(* IEC 61131-3 sources: Test-Git_ESME26/TestProgettoESME_26.fbsproj/PacDriveLib Migration/Motion/Homing, 18 files *)

(* ---- PDL_FC_ReadDriveEncoder.fn.st ---- *)
FUNCTION PDL_FC_ReadDriveEncoder: BOOL
VAR_INPUT
	i_ifDrive			: MOIN.IF_Axis;
	i_lrHomePos			: LREAL;
	i_lrAbsEncOffset	: LREAL;
	i_lrUserPeriod		: LREAL;
END_VAR
VAR_OUTPUT
	q_etDiag			: GD.ET_Diag := GD.ET_Diag.OK;
	q_etDiagExt			: PDL_ET_DiagExt := PDL_ET_DiagExt.OK;
	q_sMsg				: STRING[80];
END_VAR
VAR
	ifGetParentDevice   : DTSI.IF_GetParentDevice;
	ifDeviceAccess		: DTSI.IF_DeviceAccess;
	ifEncoderAccess		: DDI.IF_EncoderAccess;
	ifEncoder			: DDI.IF_Encoder;
	ifScalingAccess     : DMFI.IF_ScalingAccess;
	ifScaling		    : DMFI.IF_Scaling;
	xSuccess			: BOOL;
	lrEncoderPeriode:	LREAL;
	lrEncPosition:		LREAL;
	lrModuloPosition:	LREAL;
	lrHomePosition:		LREAL;
	lrTurns:			LREAL;
	lrEncoderRange:		LREAL;
	fbSetPos			: PLCO.MC_SetPosition;
END_VAR
VAR CONSTANT
	c_lrRealNull				: LREAL := 10E-12;
END_VAR

IF i_ifDrive = 0 THEN
	q_etDiag	:= GD.ET_Diag.InputParameterInvalid;
	q_etDiagExt := PDL_ET_DiagExt.DriveInvalid;
	q_sMsg		:= 'i_ifDrive - Invalid Interface';
	RETURN;
END_IF

xSuccess := __QUERYINTERFACE(i_ifDrive, ifGetParentDevice);
IF NOT xSuccess OR ifGetParentDevice = 0 THEN
	q_etDiag	:= GD.ET_Diag.InputParameterInvalid;
	q_etDiagExt := PDL_ET_DiagExt.DriveInvalid;
	q_sMsg		:= 'i_ifDrive - IF_GetParentDevice not implemented.';
	RETURN;
END_IF
ifDeviceAccess := ifGetParentDevice.GetParentDevice();

xSuccess := __QUERYINTERFACE(ifDeviceAccess,ifEncoderAccess );
IF (NOT xSuccess OR ifEncoderAccess = 0) THEN
	q_etDiag	:= GD.ET_Diag.InputParameterInvalid;
	q_etDiagExt := PDL_ET_DiagExt.DriveInvalid;
	q_sMsg		:= 'i_ifDrive - IF_Encoder not implemented.';
	RETURN;
END_IF
ifEncoder := ifEncoderAccess.Encoder;

xSuccess := __QUERYINTERFACE(ifDeviceAccess,ifScalingAccess );
IF (NOT xSuccess OR ifScalingAccess = 0) THEN
	q_etDiag	:= GD.ET_Diag.InputParameterInvalid;
	q_etDiagExt := PDL_ET_DiagExt.DriveInvalid;
	q_sMsg		:= 'i_ifDrive - IF_Scaling not implemented.';
	RETURN;
END_IF
ifScaling := ifScalingAccess.Scaling;
// Allgemeine Berehcnung ohne unterscheidung des Gebertyps			30.09.2009/ck
lrEncoderRange := ifEncoder.Revolutions;
IF (ABS(lrEncoderRange) < 1.0E-3) THEN
	q_etDiag	:= GD.ET_Diag.DriveConditionInvalid;
	q_etDiagExt := PDL_ET_DiagExt.DriveEncoderInvalid;
	q_sMsg		:= '';
	RETURN;
ELSE
	lrEncoderPeriode := lrEncoderRange * ifScaling.PositionResolution * TO_LREAL(ifScaling.GearIn) / TO_LREAL(ifScaling.GearOut);
END_IF

IF (i_lrUserPeriod < 0.0) THEN
	q_etDiag	:= GD.ET_Diag.InputParameterInvalid;
	q_etDiagExt := PDL_ET_DiagExt.UserPeriodRange;
	q_sMsg		:= '0.0 <= i_lrUserPeriod';

ELSIF (i_lrUserPeriod < c_lrRealNull) AND
	( (i_lrAbsEncOffset < c_lrRealNull) OR (i_lrAbsEncOffset > (lrEncoderPeriode - c_lrRealNull)) ) THEN
	q_etDiag	:= GD.ET_Diag.InputParameterInvalid;
	q_etDiagExt := PDL_ET_DiagExt.AbsEncOffsetRange;
	q_sMsg		:= STANDARD.CONCAT('0.0 < i_lrAbsEncOffset <= ', SE_CTBX.FC_LrealToString(i_sFormat := '#0.00', i_lrInput := lrEncoderPeriode - c_lrRealNull));

(* Check if UserPeriode fits into EncoderPeriode *)
ELSIF(i_lrUserPeriod > c_lrRealNull) AND
		(ABS(lrEncoderPeriode/i_lrUserPeriod - TRUNC_INT(lrEncoderPeriode / i_lrUserPeriod)) > c_lrRealNull ) THEN
	q_etDiag	:= GD.ET_Diag.InputParameterInvalid;
	q_etDiagExt := PDL_ET_DiagExt.UserPeriodRange;
	q_sMsg		:= STANDARD.CONCAT('i_lrUserPeriod has to be a divsior of ', SE_CTBX.FC_LrealToString(i_sFormat := '#0.00', i_lrInput := lrEncoderPeriode));

ELSE

	IF NOT ifScaling.InvertDirection THEN				(* motor direction right (true) *)
		lrEncPosition := ifEncoder.Position;
	ELSE
		lrEncPosition := lrEncoderPeriode - ifEncoder.Position;
	END_IF

(* In a round axis, position is always within the user period *)
	IF i_lrUserPeriod > c_lrRealNull THEN
		lrHomePosition := i_lrHomePos + lrEncPosition - lrEncoderPeriode/2.0;

		lrTurns :=  TRUNC_INT(lrHomePosition / i_lrUserPeriod);
		IF lrHomePosition < 0 THEN
			lrTurns := lrTurns - 1;
		END_IF

		lrModuloPosition := lrHomePosition - lrTurns * i_lrUserPeriod;

	ELSE
		lrModuloPosition := i_lrHomePos + lrEncPosition - i_lrAbsEncOffset;
	END_IF

	fbSetPos(Axis := i_ifDrive, Position := lrModuloPosition, Relative := FALSE, Execute := TRUE);

	IF fbSetPos.Error THEN
		q_etDiag	:= GD.ET_Diag.UnexpectedProgramBehavior;
		q_etDiagExt := PDL_ET_DiagExt.UnexpectedDiagExt;
		q_sMsg		:= CONCAT('Setpos: ', TO_STRING(fbSetPos.ErrorId));
	END_IF
END_IF

(* ---- PDL_FC_RestoreAxisPosition.fn.st ---- *)
FUNCTION PDL_FC_RestoreAxisPosition : BOOL
VAR_INPUT
	i_ifDrive           : MOIN.IF_Axis;
	i_lrUserPeriod      : LREAL;
	i_lrRestoreWindow   : LREAL;
	i_stRestorePosition : PDL_ST_AxisRestorePosition;
END_VAR
VAR_OUTPUT
	q_etDiag    : GD.ET_Diag     := GD.ET_Diag.OK;
	q_etDiagExt : PDL_ET_DiagExt := PDL_ET_DiagExt.OK;
	q_sMsg      : STRING[80];
END_VAR
VAR
	xSuccess            : BOOL;
	lrEncMaxPos         : LREAL;
	lrEncDiff           : LREAL;
	lrCalcAxisPos       : LREAL;
	dinPeriode          : DINT;
	diSercosState       : DINT;
	lrEncPos            : LREAL;
	lrAxisPosition      : LREAL;
	lrEncPosition       : LREAL;
	lrCheckSum          : LREAL;
	lrAxisEncPosition   : LREAL;
	lrAxisEncPosition2  : LREAL;
	diAxisGearIn        : DINT;
	diAxisGearOut       : DINT;
	lrAxisFeedConstant  : LREAL;
	diCount             : DINT;
	lrEncoderRange      : LREAL;
	ifScalingAccess     : DMFI.IF_ScalingAccess;
	ifScaling           : DMFI.IF_Scaling;
	ifGetParentDevice   : DTSI.IF_GetParentDevice;
	ifDeviceAccess      : DTSI.IF_DeviceAccess;
	ifEncoderAccess     : DDI.IF_EncoderAccess;
	ifEncoder           : DDI.IF_Encoder;
	fbSetPos            : PLCO.MC_SetPosition;
	xAxisDirection      : BOOL;

END_VAR
VAR CONSTANT
	c_lrDelta : LREAL := 0.01;
END_VAR

IF i_ifDrive = 0 THEN
	q_etDiag	:= GD.ET_Diag.InputParameterInvalid;
	q_etDiagExt := PDL_ET_DiagExt.DriveInvalid;
	q_sMsg		:= 'i_ifDrive - Invalid Interface';
	RETURN;
END_IF

xSuccess := __QUERYINTERFACE(i_ifDrive, ifGetParentDevice);
IF NOT xSuccess OR ifGetParentDevice = 0 THEN
	q_etDiag	:= GD.ET_Diag.InputParameterInvalid;
	q_etDiagExt := PDL_ET_DiagExt.DriveInvalid;
	q_sMsg		:= 'i_ifDrive - IF_GetParentDevice not implemented.';
	RETURN;
END_IF

ifDeviceAccess := ifGetParentDevice.GetParentDevice();

xSuccess := __QUERYINTERFACE(ifDeviceAccess,ifScalingAccess );
IF (NOT xSuccess OR ifScalingAccess = 0) THEN
	q_etDiag	:= GD.ET_Diag.InputParameterInvalid;
	q_etDiagExt := PDL_ET_DiagExt.DriveInvalid;
	q_sMsg		:= 'i_ifDrive - IF_Scaling not implemented.';
	RETURN;
END_IF
ifScaling := ifScalingAccess.Scaling;

xSuccess := __QUERYINTERFACE(ifDeviceAccess,ifEncoderAccess );
IF (NOT xSuccess OR ifEncoderAccess = 0) THEN
	q_etDiag	:= GD.ET_Diag.InputParameterInvalid;
	q_etDiagExt := PDL_ET_DiagExt.DriveInvalid;
	q_sMsg		:= 'i_ifDrive - IF_Encoder not implemented.';
	RETURN;
END_IF
ifEncoder := ifEncoderAccess.Encoder;

(*--------------------------------------------------------------------------------------------------------------------------------------------------*)
(* read values *)
(*--------------------------------------------------------------------------------------------------------------------------------------------------*)
	lrAxisPosition := i_stRestorePosition.lrAxisPosition;
	lrEncPosition := i_stRestorePosition.lrEncPosition;
	lrCheckSum := i_stRestorePosition.lrCheckSum;

	IF (((lrAxisPosition + lrEncPosition + c_lrDelta) < lrCheckSum) OR
		((lrAxisPosition + lrEncPosition - c_lrDelta) > lrCheckSum)) THEN

		q_etDiag	:= GD.ET_Diag.InputParameterInvalid;
		q_etDiagExt := PDL_ET_DiagExt.CheckSumInvalid;
		q_sMsg		:= '';
		RETURN;
	END_IF

(*--------------------------------------------------------------------------------------------------------------------------------------------------*)
(* Check Sercos state and read values *)
(*--------------------------------------------------------------------------------------------------------------------------------------------------*)
FOR diCount := 1 TO 3 DO

	diSercosState := FC_GetSercosState();
	IF diSercosState = 4 THEN
		lrAxisEncPosition := ifEncoder.Position;
		diAxisGearIn := TO_DINT(ifScaling.GearIn);
		diAxisGearOut := TO_DINT(ifScaling.GearOut);
		lrAxisFeedConstant := ifScaling.PositionResolution;
		xAxisDirection := NOT ifScaling.InvertDirection;
	ELSE
		q_etDiag	:= GD.ET_Diag.SercosConditionInvalid;
		q_etDiagExt := PDL_ET_DiagExt.SercosNotInPhaseFour;
		q_sMsg		:= '';
		RETURN;
	END_IF

(*--------------------------------------------------------------------------------------------------------------------------------------------------*)
(* Berechnung der maximale Encoder Position *)
(*--------------------------------------------------------------------------------------------------------------------------------------------------*)

	// Allgemeine Berechnung ohne Unterscheidung des Gebertyps
	lrEncoderRange := ifEncoder.Revolutions;
	IF (ABS(lrEncoderRange) < 1.0E-3) THEN
		q_etDiag	:= GD.ET_Diag.DriveConditionInvalid;
		q_etDiagExt := PDL_ET_DiagExt.DriveEncoderInvalid;
		q_sMsg		:= '';
		RETURN;
	ELSE
		lrEncMaxPos := lrEncoderRange * lrAxisFeedConstant * TO_LREAL(diAxisGearIn) / TO_LREAL(diAxisGearOut);
	END_IF

(*--------------------------------------------------------------------------------------------------------------------------------------------------*)
(* Differenz der Geberposition *)
(*--------------------------------------------------------------------------------------------------------------------------------------------------*)
	IF xAxisDirection THEN		(* +++ Rechtslauf +++ *)
		lrEncDiff := lrAxisEncPosition - lrEncPosition;
		IF lrEncDiff > lrEncMaxPos/2 THEN
			lrEncPos := lrAxisEncPosition - lrEncMaxPos;
			lrEncDiff := lrEncDiff - lrEncMaxPos;
		ELSIF lrEncDiff < -lrEncMaxPos/2 THEN
			lrEncPos := lrAxisEncPosition + lrEncMaxPos;
			lrEncDiff := lrEncDiff + lrEncMaxPos ;
		ELSE
			lrEncPos := lrAxisEncPosition;
		END_IF
		lrCalcAxisPos := lrEncPos - lrEncPosition + lrAxisPosition;

	ELSE						(* +++ Linkslauf +++ *)
		lrEncDiff:=  lrEncPosition - lrAxisEncPosition;	(*  lrEncMaxPos - lrAxisEncPosition
																 - (lrEncMaxPos- lrEncPos_Retain) *)
		IF lrEncDiff > lrEncMaxPos/2 THEN
			lrEncPos :=  - lrAxisEncPosition;				(* lrEncMaxPos - lrAxisEncPosition - lrEncMaxPos *)
			lrEncDiff := lrEncDiff - lrEncMaxPos;
		ELSIF lrEncDiff < -lrEncMaxPos/2 THEN
			lrEncPos := 2*lrEncMaxPos - lrAxisEncPosition;	(* lrEncMaxPos - lrAxisEncPosition + lrEncMaxPos *)
			lrEncDiff := lrEncDiff + lrEncMaxPos ;
		ELSE
			lrEncPos := lrEncMaxPos - lrAxisEncPosition;
		END_IF
		lrCalcAxisPos := lrEncPos -  (lrEncMaxPos - lrEncPosition) + lrAxisPosition;
	END_IF

(*--------------------------------------------------------------------------------------------------------------------------------------------------*)
(* check if in Window *)
(*--------------------------------------------------------------------------------------------------------------------------------------------------*)
	IF ABS(lrEncDiff) > ABS(i_lrRestoreWindow) THEN	(* Maximale Abweichung prüfen *)
		q_etDiag	:= GD.ET_Diag.DriveConditionInvalid;
		q_etDiagExt := PDL_ET_DiagExt.OutOfRestoreWindow;
		q_sMsg		:= '';
		RETURN;

(*--------------------------------------------------------------------------------------------------------------------------------------------------*)
(* Set axis position *)
(*--------------------------------------------------------------------------------------------------------------------------------------------------*)
	ELSE
		IF i_lrUserPeriod > 0 THEN
			dinPeriode:=TRUNC_INT(lrCalcAxisPos / i_lrUserPeriod );
			IF lrCalcAxisPos < 0.0 THEN
				dinPeriode:= dinPeriode - 1;
			END_IF
			lrCalcAxisPos:= lrCalcAxisPos - (dinPeriode * i_lrUserPeriod);
		END_IF

		fbSetPos(Axis := i_ifDrive, Position := lrCalcAxisPos, Relative := FALSE, Execute := TRUE);
		IF fbSetPos.Error THEN
			q_etDiag	:= GD.ET_Diag.UnexpectedProgramBehavior;
			q_etDiagExt := PDL_ET_DiagExt.UnexpectedFeedback;
			q_sMsg		:= CONCAT('Setpos: ', PLCO.FC_EtResultToString(fbSetPos.ErrorId));
		END_IF

	END_IF

	(* read again to make shure, that there was no interrupt through the Sercos *)
	lrAxisEncPosition2 :=  ifEncoder.Position;
	IF ABS(	lrAxisEncPosition - lrAxisEncPosition2) < c_lrDelta THEN
		RETURN;
	END_IF
END_FOR

q_etDiag	:= GD.ET_Diag.DriveConditionInvalid;
q_etDiagExt := PDL_ET_DiagExt.RestoreInterrupted;
q_sMsg		:= '';

(* ---- PDL_FC_SaveAxisPosition.fn.st ---- *)
FUNCTION PDL_FC_SaveAxisPosition : BOOL
VAR_INPUT
	i_etPosType : PDL_ET_PosType;
	i_ifDrive   : MOIN.IF_Axis;
END_VAR

VAR_IN_OUT
	iq_stRestorePosition : PDL_ST_AxisRestorePosition;
END_VAR

VAR_OUTPUT
	q_etDiag    : GD.ET_Diag     := GD.ET_Diag.OK;
	q_etDiagExt : PDL_ET_DiagExt := PDL_ET_DiagExt.OK;
	q_sMsg      : STRING[80];
END_VAR

VAR
	etSercosState       : SMI.ET_SercosState;
	xSuccess            : BOOL;
	lrAxisPosition      : LREAL;
	lrEncPosition       : LREAL;
	lrAxisPosition2     : LREAL;
	lrEncPosition2      : LREAL;
	diCount             : DINT;
	ifDriveAccess       : DMFI.IF_DriveAccess;
	ifDrive             : DMFI.IF_Drive;
	ifEncoderAccess     : DDI.IF_EncoderAccess;
	ifEncoder           : DDI.IF_Encoder;
	ifGetParentDevice   : DTSI.IF_GetParentDevice;
	ifDeviceAccess      : DTSI.IF_DeviceAccess;

END_VAR

VAR CONSTANT
	c_lrDelta : LREAL := 0.01;

END_VAR

IF i_ifDrive = 0 THEN
	q_etDiag    := GD.ET_Diag.InputParameterInvalid;
	q_etDiagExt := PDL_ET_DiagExt.DriveInvalid;
	q_sMsg      := 'i_ifDrive - Invalid Interface';
	RETURN;
END_IF

xSuccess := __QUERYINTERFACE(i_ifDrive, ifGetParentDevice);
IF NOT xSuccess OR ifGetParentDevice = 0 THEN
	q_etDiag    := GD.ET_Diag.InputParameterInvalid;
	q_etDiagExt := PDL_ET_DiagExt.DriveInvalid;
	q_sMsg      := 'i_ifDrive - IF_GetParentDevice not implemented.';
	RETURN;
END_IF
ifDeviceAccess := ifGetParentDevice.GetParentDevice();

xSuccess := __QUERYINTERFACE(ifDeviceAccess, ifDriveAccess);
IF (NOT xSuccess OR ifDriveAccess = 0) THEN
	q_etDiag    := GD.ET_Diag.InputParameterInvalid;
	q_etDiagExt := PDL_ET_DiagExt.DriveInvalid;
	q_sMsg      := 'i_ifDrive - IF_Drive not implemented.';
	RETURN;
END_IF
ifDrive := ifDriveAccess.Drive;

xSuccess := __QUERYINTERFACE(ifDeviceAccess, ifEncoderAccess);
IF (NOT xSuccess OR ifEncoderAccess = 0) THEN
	q_etDiag    := GD.ET_Diag.InputParameterInvalid;
	q_etDiagExt := PDL_ET_DiagExt.DriveInvalid;
	q_sMsg      := 'i_ifDrive - IF_Encoder not implemented.';
	RETURN;
END_IF
ifEncoder := ifEncoderAccess.Encoder;

FOR diCount := 1 TO 3 DO

	etSercosState := FC_GetSercosState();
	IF etSercosState = SMI.ET_SercosState.Phase4 THEN

		(* first read of AxisPos and EncoderPos *)
		CASE i_etPosType OF
			PDL_ET_PosType.Position:
				lrAxisPosition := ifDrive.ActualPosition;
			PDL_ET_PosType.RefPosition:
				lrAxisPosition := i_ifDrive.RefPosition;
			PDL_ET_PosType.MechPosition:
				lrAxisPosition := ifDrive.ActualPosition;
			PDL_ET_PosType.MechRefPosition:
				lrAxisPosition := i_ifDrive.RefPosition;
			ELSE
				lrAxisPosition := i_ifDrive.RefPosition;
		END_CASE

		lrEncPosition := ifEncoder.Position;

		(* second read of AxisPos and EncoderPos *)
		CASE i_etPosType OF
			PDL_ET_PosType.Position:
				lrAxisPosition2 := ifDrive.ActualPosition;
			PDL_ET_PosType.RefPosition:
				lrAxisPosition2 := i_ifDrive.RefPosition;
			PDL_ET_PosType.MechPosition:
				lrAxisPosition2 := ifDrive.ActualPosition;
			PDL_ET_PosType.MechRefPosition:
				lrAxisPosition2 := i_ifDrive.RefPosition;
			ELSE
				lrAxisPosition2 := i_ifDrive.RefPosition;
		END_CASE

		lrEncPosition2 := ifEncoder.Position;

	ELSE
		q_etDiag    := GD.ET_Diag.SercosConditionInvalid;
		q_etDiagExt := PDL_ET_DiagExt.SercosNotInPhaseFour;
		q_sMsg      := '';
		RETURN;
	END_IF

	IF (ABS(lrEncPosition - lrEncPosition2) < c_lrDelta) AND (ABS(lrAxisPosition - lrAxisPosition2) < c_lrDelta) THEN
		EXIT;
	END_IF
END_FOR

etSercosState := FC_GetSercosState();
IF (etSercosState = SMI.ET_SercosState.Phase4) AND (diCount <= 3) THEN
	iq_stRestorePosition.lrAxisPosition := lrAxisPosition2;
	iq_stRestorePosition.lrEncPosition  := lrEncPosition2;
	iq_stRestorePosition.lrCheckSum     := lrAxisPosition2 + lrEncPosition2;
ELSE
	q_etDiag    := GD.ET_Diag.SercosConditionInvalid;
	q_etDiagExt := PDL_ET_DiagExt.SercosNotInPhaseFour;
	q_sMsg      := '';
END_IF

(* ---- PDL_FB_Home.fb.st ---- *)
FUNCTION_BLOCK PDL_FB_Home
VAR_INPUT
	i_xEnable     : BOOL;
	i_etMode      : PDL_ET_HomeMode := PDL_ET_HomeMode.SetPosAxisAndLogEncoderPosition;
	i_ifDrive     : Moin.IF_Axis;
	i_xHwLimitNeg : BOOL;
	i_xHwLimitPos : BOOL;
	i_xStart      : BOOL;
END_VAR
VAR_OUTPUT
	q_xActive                  : BOOL;
	q_xReady                   : BOOL;
	q_etDiag                   : GD.ET_Diag := GD.ET_Diag.Ok;
	q_etDiagExt                : PDL_ET_DiagExt := PDL_ET_DiagExt.Disabled;
	q_sMsg                     : STRING[80];
	q_xDisableDrive            : BOOL  := FALSE;
	q_xMotionInstructionActive : BOOL;
	q_lrPosition               : LREAL := 0.0;
	q_lrEncoderPosition        : LREAL := 0.0;
	q_xHomeOk                  : BOOL;
END_VAR
VAR
	stSensor_loc           : PDL_ST_HomeIn;
	stLimitSwitch_loc      : PDL_ST_HomeLimitSwitch;
	stMoveOnPos_loc        : PDL_ST_HomeMoveOnPos;
	stSetPos_loc           : PDL_ST_HomeSetPos;
	stTorque_loc           : PDL_ST_HomeTorque;
	stForce_loc            : PDL_ST_HomeForce;
	stTouchProbe_loc       : PDL_ST_HomeTp;
	stWritePos_loc         : PDL_ST_HomeWritePos;
	stReducedVelocity_loc  : PDL_ST_ReducedVelocity;
	xEnableFlag            : BOOL;
	etHomeState            : PDL_ET_HomeState;
	etHomeOpMode           : PDL_ET_HomeOpMode;
	xStartFlag             : BOOL;
	xStartHomeIn           : BOOL;
	fbHomeTP               : PDL_FB_HomeTp;
	fbHomeIn               : PDL_FB_HomeIn;
	fbHomeLS               : PDL_FB_HomeLimitSwitch;
	fbHomeTorque           : PDL_FB_HomeTorque;
	fbHomeForce            : PDL_FB_HomeForce;
	fbVarioPosJerk         : PDL_FB_VarioPosJerk;
	fbHomeAbs              : PDL_FB_HomeAbs;
	fbSetpos               : PDL_FB_HomeSetpos;
	etHomeTpMode           : PDL_ET_HomeTpMode;
	etHomeInMode           : PDL_ET_HomeInMode;
	etHomeLimitSwitchMode  : PDL_ET_HomeLimitSwitchMode;
	etHomeTorqueMode       : PDL_ET_HomeTorqueMode;
	etHomeForceMode        : PDL_ET_HomeForceMode;
	etHomeSetPosMode       : PDL_ET_HomeSetPosMode;
	xSuccess               : BOOL;
	xFbEnable              : BOOL;
	xFbActive              : BOOL;
	lrUsedVelocity         : LREAL;
	lrLowVelocity          : LREAL;
	etDiagBuffer           : GD.ET_Diag;
	sTempMsg               : STRING[80] := '';
	xFbHomeOk              : BOOL;
	lrPositionOpmMoveOnPos : LREAL;
	xDetectSetPosHomeOnPos : BOOL;
	fbLoggerPoint          : APL.FB_LoggerPoint;
	xControllerStop        : BOOL;
	fbTrigStop              : Standard.R_TRIG;
	fbSetPosIntern         : PLCO.MC_SetPosition;
	ifGetParentDevice      : DTSI.IF_GetParentDevice;
	ifDeviceAccess         : DTSI.IF_DeviceAccess;
	ifDriveAccess          : DMFI.IF_DriveAccess;
	ifDrive                : DMFI.IF_Drive;

	xInitReducedVel : BOOL;
END_VAR

(* ------------------------------------------------------------------------------------------------------------------------------------------------------*)
(* Wait for Enable *)
(* ------------------------------------------------------------------------------------------------------------------------------------------------------*)
IF i_xEnable AND NOT xEnableflag THEN (*  Input action by rising edge of enable *)
	xEnableFlag := TRUE;
	THIS^.fbLoggerPoint.AddLogEntry(
		i_etLogLevel := APL.ET_LogLevel.UserAction,
		i_etDiag     := q_etDiag,
		i_udiDiagExt := q_etDiagExt,
		i_sMessage   := 'enable function block',
		q_etDiag     =>,
		q_etDiagExt  =>
	);
	q_xActive                  := TRUE;
	q_xReady                   := FALSE;
	q_xDisableDrive            := FALSE;
	q_xMotionInstructionActive := FALSE;

	xFbEnable  := FALSE;
	xStartFlag := FALSE;
	q_xReady   := TRUE;
	SetDiagOutput(i_etDiag := GD.ET_Diag.OK, i_etDiagExt := PDL_ET_DiagExt.WaitForStart, i_sMsg := '');
	etHomeState := PDL_ET_HomeState.WaitForStart;

ELSIF NOT i_xEnable AND xEnableflag THEN (* Input action by falling edge of enable *)
	xEnableFlag := FALSE;
	THIS^.fbLoggerPoint.AddLogEntry(
		i_etLogLevel := APL.ET_LogLevel.UserAction,
		i_etDiag     := q_etDiag,
		i_udiDiagExt := q_etDiagExt,
		i_sMessage   := 'disable function block',
		q_etDiag     =>,
		q_etDiagExt  =>
	);
	q_xReady  := FALSE;
	xFbEnable := FALSE;
	SetDiagOutput(i_etDiag := GD.ET_Diag.Ok, i_etDiagExt := PDL_ET_DiagExt.WaitUntilDisabled, i_sMsg := '');
	etHomeState := PDL_ET_HomeState.WaitUntilDisabled; (* Wait until disabled *)
END_IF

IF NOT i_xStart AND xStartFlag THEN (* allways accept the falling edge in i_xStart *)
	xStartFlag := FALSE; (* make no difference for the fbs called inside, because their start ist fixed to TRUE *)
END_IF

(* Continuous Checks at Enable *)
IF i_xEnable THEN
	(* Check HW-Limits in Pos-Mode because FB_VarioPosJerk has no HW-Limit-Inputs *)
	IF
		(etHomeOpMode = PDL_ET_HomeOpMode.Torque OR etHomeOpMode = PDL_ET_HomeOpMode.Force OR etHomeOpMode = PDL_ET_HomeOpMode.MoveOnPos) AND
		(i_xHwLimitNeg OR i_xHwLimitPos)
	THEN
		IF i_xHwLimitNeg THEN
			SetDiagOutput(i_etDiag := GD.ET_Diag.LimitReached, i_etDiagExt := PDL_ET_DiagExt.HwLimitNegReached, i_sMsg := '');
		ELSIF i_xHwLimitPos THEN
			SetDiagOutput(i_etDiag := GD.ET_Diag.LimitReached, i_etDiagExt := PDL_ET_DiagExt.HwLimitPosReached, i_sMsg := '');
		END_IF
	END_IF
	(* Check ReducedVelocity *)
	IF stReducedVelocity_loc.i_xEnableReducedVelocity THEN
		IF NOT xInitReducedVel THEN
			xInitReducedVel := TRUE;
			(* Check Interfaces *)
			xSuccess := __QUERYINTERFACE(i_ifDrive, ifGetParentDevice);
			IF NOT xSuccess OR ifGetParentDevice = 0 THEN
				SetDiagOutput(
					i_etDiag    := GD.ET_Diag.InputParameterInvalid,
					i_etDiagExt := PDL_ET_DiagExt.DriveInvalid,
					i_sMsg      := 'i_ifDrive - IF_GetParentDevice not implemented.'
				);
			END_IF
			ifDeviceAccess := ifGetParentDevice.GetParentDevice();

			xSuccess := __QUERYINTERFACE(ifDeviceAccess, ifDriveAccess);
			IF (NOT xSuccess OR ifDriveAccess = 0) THEN
				SetDiagOutput(
					i_etDiag    := GD.ET_Diag.InputParameterInvalid,
					i_etDiagExt := PDL_ET_DiagExt.DriveInvalid,
					i_sMsg      := 'i_ifDrive - IF_Drive not implemented.'
				);
			END_IF
			ifDrive := ifDriveAccess.Drive;
		END_IF

		IF stReducedVelocity_loc.i_lrMaxReducedVelocity <= 0 THEN
			SetDiagOutput(
				i_etDiag    := GD.ET_Diag.InputParameterInvalid,
				i_etDiagExt := PDL_ET_DiagExt.ReducedVelocityRange,
				i_sMsg      := 'lrMaxReducedVelocity <= 0'
			);
		END_IF
		IF stReducedVelocity_loc.i_lrReducedVelocityCheckFactor < 1.0 THEN
			SetDiagOutput(
				i_etDiag    := GD.ET_Diag.InputParameterInvalid,
				i_etDiagExt := PDL_ET_DiagExt.ReducedVelocityFactorRange,
				i_sMsg      := 'i_lrReducedVelocityCheckFactor < 1'
			);
		END_IF
		IF ifDrive <> 0 THEN
			IF
				ABS(ifDrive.ActualPosition) > ABS(stReducedVelocity_loc.i_lrMaxReducedVelocity * stReducedVelocity_loc.i_lrReducedVelocityCheckFactor)
			THEN
				SetDiagOutput(i_etDiag := GD.ET_Diag.LimitReached, i_etDiagExt := PDL_ET_DiagExt.ReducedVelocityLimit, i_sMsg := '');
			END_IF
		END_IF
	ELSE
		xInitReducedVel := FALSE;
	END_IF
END_IF

(*Statemachine*)
//etHomeState is also changed in SetDiagOutput and Diag-Translations at END of HomingOpModes-Blocks in FB_Home AS-Structure
CASE etHomeState OF
	(* ------------------------------------------------------------------------------------------------------------------------------------------------------*)
	PDL_ET_HomeState.ExceptionOrIdle: (* Idle or Error *)
		(* ------------------------------------------------------------------------------------------------------------------------------------------------------*)
		;

		(* ------------------------------------------------------------------------------------------------------------------------------------------------------*)
	PDL_ET_HomeState.WaitForStart: (* Wait for Start *)
		(* ------------------------------------------------------------------------------------------------------------------------------------------------------*)
		IF i_xStart AND NOT xStartFlag THEN
			xStartFlag := TRUE;
			THIS^.fbLoggerPoint.AddLogEntry(
				i_etLogLevel := APL.ET_LogLevel.UserAction,
				i_etDiag     := q_etDiag,
				i_udiDiagExt := q_etDiagExt,
				i_sMessage   := 'start function block',
				q_etDiag     =>,
				q_etDiagExt  =>
			);
			q_xHomeOK := FALSE;
			sTempMsg  := '';
			IF
				i_etMode = PDL_ET_HomeMode.PosDirectionPosEdgeTp OR
				i_etMode = PDL_ET_HomeMode.NegDirectionPosEdgeTp OR
				i_etMode = PDL_ET_HomeMode.NegDirectionNegEdgeTp OR
				i_etMode = PDL_ET_HomeMode.PosDirectionNegEdgeTp
			THEN (* HomeTP *)

				etHomeOpMode := PDL_ET_HomeOpMode.TouchProbe;
				CASE i_etMode OF
					PDL_ET_HomeMode.PosDirectionPosEdgeTp:
						etHomeTpMode := PDL_ET_HomeTpMode.PosDirectionPosEdgeTp;
					PDL_ET_HomeMode.NegDirectionPosEdgeTp:
						etHomeTpMode := PDL_ET_HomeTpMode.NegDirectionPosEdgeTp;
					PDL_ET_HomeMode.NegDirectionNegEdgeTp:
						etHomeTpMode := PDL_ET_HomeTpMode.NegDirectionNegEdgeTp;
					PDL_ET_HomeMode.PosDirectionNegEdgeTp:
						etHomeTpMode := PDL_ET_HomeTpMode.PosDirectionNegEdgeTp;
				END_CASE
				xFbEnable := TRUE;
				sTempMsg  := 'HomeTP';
				DriveAndLencCheck();
				THIS^.fbHomeTP.RegisterLoggerPoint(i_ifParent := THIS^.fbLoggerPoint, i_sName := 'HomeTp', q_etDiag =>, q_etDiagExt => );
				(* HomeIN *)
			ELSIF
				i_etMode = PDL_ET_HomeMode.PosDirectionPosEdgeSensor OR
				i_etMode = PDL_ET_HomeMode.NegDirectionPosEdgeSensor OR
				i_etMode = PDL_ET_HomeMode.NegDirectionNegEdgeSensor OR
				i_etMode = PDL_ET_HomeMode.PosDirectionNegEdgeSensor
			THEN

				etHomeOpMode := PDL_ET_HomeOpMode.Sensor;
				CASE i_etMode OF
					PDL_ET_HomeMode.PosDirectionPosEdgeSensor:
						etHomeInMode := PDL_ET_HomeInMode.PosDirectionPosEdgeSensor;
					PDL_ET_HomeMode.NegDirectionPosEdgeSensor:
						etHomeInMode := PDL_ET_HomeInMode.NegDirectionPosEdgeSensor;
					PDL_ET_HomeMode.NegDirectionNegEdgeSensor:
						etHomeInMode := PDL_ET_HomeInMode.NegDirectionNegEdgeSensor;
					PDL_ET_HomeMode.PosDirectionNegEdgeSensor:
						etHomeInMode := PDL_ET_HomeInMode.PosDirectionNegEdgeSensor;
				END_CASE
				xStartHomeIn := FALSE;
				xFbEnable    := TRUE;
				sTempMsg     := 'HomeIn';
				DriveAndLencCheck();
				THIS^.fbHomeIn.RegisterLoggerPoint(i_ifParent := THIS^.fbLoggerPoint, i_sName := 'HomeIn', q_etDiag =>, q_etDiagExt => );
				(* HomeLS *)
			ELSIF
				i_etMode = PDL_ET_HomeMode.PosDirectionPosEdgeHWLimitPos OR
				i_etMode = PDL_ET_HomeMode.NegDirectionPosEdgeHWLimitNeg OR
				i_etMode = PDL_ET_HomeMode.NegDirectionNegEdgeHWLimitNeg OR
				i_etMode = PDL_ET_HomeMode.PosDirectionNegEdgeHWLimitPos
			THEN

				etHomeOpMode := PDL_ET_HomeOpMode.LimitSwitch;
				CASE i_etMode OF
					PDL_ET_HomeMode.PosDirectionPosEdgeHWLimitPos:
						etHomeLimitSwitchMode := PDL_ET_HomeLimitSwitchMode.PosDirectionPosEdgeHWLimitPos;
					PDL_ET_HomeMode.NegDirectionPosEdgeHWLimitNeg:
						etHomeLimitSwitchMode := PDL_ET_HomeLimitSwitchMode.NegDirectionPosEdgeHWLimitNeg;
					PDL_ET_HomeMode.NegDirectionNegEdgeHWLimitNeg:
						etHomeLimitSwitchMode := PDL_ET_HomeLimitSwitchMode.NegDirectionNegEdgeHWLimitNeg;
					PDL_ET_HomeMode.PosDirectionNegEdgeHWLimitPos:
						etHomeLimitSwitchMode := PDL_ET_HomeLimitSwitchMode.PosDirectionNegEdgeHWLimitPos;
				END_CASE
				xFbEnable := TRUE;
				sTempMsg  := 'HomeLS';
				DriveAndLencCheck();
				THIS^.fbHomeLS.RegisterLoggerPoint(i_ifParent := THIS^.fbLoggerPoint, i_sName := 'HomeLimitSwitch', q_etDiag =>, q_etDiagExt => );
				(* HomeTorque *)
			ELSIF i_etMode = PDL_ET_HomeMode.PosDirectionMaxTorque OR i_etMode = PDL_ET_HomeMode.NegDirectionMaxTorque THEN

				etHomeOpMode := PDL_ET_HomeOpMode.Torque;
				CASE i_etMode OF
					PDL_ET_HomeMode.PosDirectionMaxTorque:
						etHomeTorqueMode := PDL_ET_HomeTorqueMode.PosDirectionMaxTorque;
					PDL_ET_HomeMode.NegDirectionMaxTorque:
						etHomeTorqueMode := PDL_ET_HomeTorqueMode.NegDirectionMaxTorque;
				END_CASE
				xFbEnable := TRUE;
				sTempMsg  := 'HomeTorque';
				DriveAndLencCheck();
				THIS^.fbHomeTorque.RegisterLoggerPoint(i_ifParent := THIS^.fbLoggerPoint, i_sName := 'HomeTorque', q_etDiag =>, q_etDiagExt => );

			ELSIF i_etMode = PDL_ET_HomeMode.PosDirectionMaxForce OR i_etMode = PDL_ET_HomeMode.NegDirectionMaxForce THEN

				SetDiagOutput(
					i_etDiag    := GD.ET_Diag.InputParameterInvalid,
					i_etDiagExt := PDL_ET_DiagExt.UnknownMode,
					i_sMsg      := concat('HomeMode not yet supported', TO_STRING(i_etMode))
				);
				RETURN;

			ELSIF i_etMode = PDL_ET_HomeMode.MoveOnPosAbs THEN (* Home move on Pos *)

				etHomeOpMode := PDL_ET_HomeOpMode.MoveOnPos;
				IF stMoveOnPos_loc.i_lrPeriod > 0 AND stMoveOnPos_loc.i_xRotativeSystem THEN
					lrPositionOpmMoveOnPos :=
						MATH.fmod(lrX := (stMoveOnPos_loc.i_lrTarget - i_ifDrive.lrPosition), lrM := stMoveOnPos_loc.i_lrPeriod);
					IF lrPositionOpmMoveOnPos > stMoveOnPos_loc.i_lrPeriod / 2 THEN
						lrPositionOpmMoveOnPos := lrPositionOpmMoveOnPos - stMoveOnPos_loc.i_lrPeriod;
					END_IF
					IF lrPositionOpmMoveOnPos < -stMoveOnPos_loc.i_lrPeriod / 2 THEN
						lrPositionOpmMoveOnPos := lrPositionOpmMoveOnPos + stMoveOnPos_loc.i_lrPeriod;
					END_IF
				ELSE
					lrPositionOpmMoveOnPos := stMoveOnPos_loc.i_lrTarget;
				END_IF

				xControllerStop := FALSE;

				fbVarioPosJerk(i_ifDrive := i_ifDrive, i_xEnable := FALSE, i_xStart := FALSE, i_xStop := FALSE);
				xFbEnable := TRUE;
				sTempMsg  := 'MoveOnPosAbs';
				DriveAndLencCheck();
				THIS^.fbVarioPosJerk.RegisterLoggerPoint(i_ifParent := THIS^.fbLoggerPoint, i_sName := 'MoveOnPosAbs', q_etDiag =>, q_etDiagExt => );

			ELSIF i_etMode = PDL_ET_HomeMode.WriteAxisEncoder THEN (* HomeAbs *)

				etHomeOpMode := PDL_ET_HomeOpMode.WritePos;
				xFbEnable    := TRUE;
				sTempMsg     := 'WritePos';
				DriveAndLencCheck(); (* HomeSetPos *)
				THIS^.fbHomeAbs.RegisterLoggerPoint(i_ifParent := THIS^.fbLoggerPoint, i_sName := 'HomeAbs', q_etDiag =>, q_etDiagExt => );

			ELSIF
				i_etMode = PDL_ET_HomeMode.SetPosAxisPosition OR
				i_etMode = PDL_ET_HomeMode.SetPosLogEncoderPosition OR
				i_etMode = PDL_ET_HomeMode.SetPosAxisAndLogEncoderPosition OR
				i_etMode = PDL_ET_HomeMode.RestorePosFromAxisEncoder OR
				i_etMode = PDL_ET_HomeMode.RestorePosFromRetain
			THEN

				etHomeOpMode := PDL_ET_HomeOpMode.SetPos;
				CASE i_etMode OF
					PDL_ET_HomeMode.SetPosAxisPosition:
						etHomeSetPosMode := PDL_ET_HomeSetPosMode.SetPosAxisPosition;
					PDL_ET_HomeMode.SetPosLogEncoderPosition:
						etHomeSetPosMode := PDL_ET_HomeSetPosMode.SetPosLogEncoderPosition;
					PDL_ET_HomeMode.SetPosAxisAndLogEncoderPosition:
						etHomeSetPosMode := PDL_ET_HomeSetPosMode.SetPosAxisAndLogEncoderPosition;
					PDL_ET_HomeMode.RestorePosFromAxisEncoder:
						etHomeSetPosMode := PDL_ET_HomeSetPosMode.RestorePosFromAxisEncoder;
					PDL_ET_HomeMode.RestorePosFromRetain:
						etHomeSetPosMode := PDL_ET_HomeSetPosMode.RestorePosFromRetain;
				END_CASE
				xFbEnable := TRUE;
				sTempMsg  := 'HomeSetPos';
				DriveAndLencCheck();
				THIS^.fbSetpos.RegisterLoggerPoint(i_ifParent := THIS^.fbLoggerPoint, i_sName := 'HomeSetPos', q_etDiag =>, q_etDiagExt => );

			ELSE
				etHomeOpMode := PDL_ET_HomeOpMode.NoOp;
				SetDiagOutput(
					i_etDiag := GD.ET_Diag.InputParameterInvalid, i_etDiagExt := PDL_ET_DiagExt.UnknownMode, i_sMsg := UDINT_TO_STRING(i_etMode)
				);
			END_IF

			IF etHomeOpMode <> PDL_ET_HomeOpMode.NoOp THEN
				SetDiagOutput(i_etDiag := GD.ET_Diag.Ok, i_etDiagExt := PDL_ET_DiagExt.WaitUntilHomingDone, i_sMsg := sTempMsg);
			END_IF
			etHomeState := PDL_ET_HomeState.WaitUntilFbActive;
		END_IF

		(* ------------------------------------------------------------------------------------------------------------------------------------------------------*)
	PDL_ET_HomeState.WaitUntilFbActive: (* Wait HomeFB active *)
		(* ------------------------------------------------------------------------------------------------------------------------------------------------------*)
		THIS^.CallFb();
		IF THIS^.xFbActive THEN
			fbLoggerPoint.AddLogEntry(
				i_etLogLevel := APL.ET_LogLevel.DebugMessage,
				i_etDiag     := q_etDiag,
				i_udiDiagExt := q_etDiagExt,
				i_sMessage   := 'Start homing',
				q_etDiag     =>,
				q_etDiagExt  =>
			);
			etHomeState := PDL_ET_HomeState.WaitUntilHomeOk;
		END_IF

		(* ------------------------------------------------------------------------------------------------------------------------------------------------------*)
	PDL_ET_HomeState.WaitUntilHomeOk: (* Wait HomeOk , Check DiagExt-Codes while Execution; If Number 30 changed, see ...TranslateDiag-Methods*)
		(* ------------------------------------------------------------------------------------------------------------------------------------------------------*)
		xStartHomeIn := TRUE;
		THIS^.CallFb();
		IF (THIS^.etDiagBuffer = GD.ET_Diag.Ok) AND THIS^.xFbHomeOk THEN
			q_xHomeOK := TRUE;
			xFbEnable := FALSE;
			SetDiagOutput(i_etDiag := GD.ET_Diag.Ok, i_etDiagExt := PDL_ET_DiagExt.HomingDone, i_sMsg := sTempMsg);
			etHomeState := PDL_ET_HomeState.WaitUntilFbDisabled;
		END_IF

		(* ------------------------------------------------------------------------------------------------------------------------------------------------------*)
	PDL_ET_HomeState.WaitUntilFbDisabled: (* Wait for FB disabled*)
		(* ------------------------------------------------------------------------------------------------------------------------------------------------------*)
		THIS^.CallFb();
		IF NOT xFbActive THEN
			q_xMotionInstructionActive := FALSE;
			etHomeOpMode               := PDL_ET_HomeOpMode.NoOp;
			fbLoggerPoint.AddLogEntry(
				i_etLogLevel := APL.ET_LogLevel.StatusMessage,
				i_etDiag     := q_etDiag,
				i_udiDiagExt := q_etDiagExt,
				i_sMessage   := 'ready for start',
				q_etDiag     =>,
				q_etDiagExt  =>
			);
			etHomeState := PDL_ET_HomeState.WaitForStart;
		END_IF

		(* ------------------------------------------------------------------------------------------------------------------------------------------------------*)
	PDL_ET_HomeState.WaitUntilDisabled: (* Wait for FB disabled*)
		(* ------------------------------------------------------------------------------------------------------------------------------------------------------*)
		THIS^.CallFb();
		IF NOT xFbActive THEN
			q_xActive                  := FALSE;
			q_xDisableDrive            := FALSE;
			q_xMotionInstructionActive := FALSE;
			q_lrPosition               := 0.0;
			q_lrEncoderPosition        := 0.0;
			q_xHomeOK                  := FALSE;
			SetDiagOutput(i_etDiag := GD.ET_Diag.Ok, i_etDiagExt := PDL_ET_DiagExt.Disabled, i_sMsg := '');
			etHomeState := PDL_ET_HomeState.ExceptionOrIdle;
		END_IF
		(* ------------------------------------------------------------------------------------------------------------------------------------------------------*)
END_CASE

IF i_xEnable THEN
	(* q_xMotionInstructionActive Set or Reset *)
	IF fbHomeIn.q_xActive THEN
		q_xMotionInstructionActive := fbHomeIn.q_xMotionInstructionActive;
	ELSIF fbHomeTP.q_xActive THEN
		q_xMotionInstructionActive := fbHomeTP.q_xMotionInstructionActive;
	ELSIF fbHomeLS.q_xActive THEN
		q_xMotionInstructionActive := fbHomeLS.q_xMotionInstructionActive;
	ELSIF fbHomeTorque.q_xActive THEN
		q_xMotionInstructionActive := fbHomeTorque.q_xMotionInstructionActive;
	ELSIF fbHomeForce.q_xActive THEN
		q_xMotionInstructionActive := fbHomeForce.q_xMotionInstructionActive;
	ELSIF fbVarioPosJerk.q_xActive THEN
		q_xMotionInstructionActive := fbVarioPosJerk.q_xMotionInstructionActive;
	ELSIF fbHomeAbs.q_xActive THEN
		q_xMotionInstructionActive := fbHomeAbs.q_xActive; // set to q_xActive, because previous version of FB has set output depending on q_xActive
	ELSIF fbSetpos.q_xActive THEN
		q_xMotionInstructionActive := fbSetpos.q_xActive; // set to q_xActive, because previous version of FB has set output depending on q_xActive
	ELSE
		q_xMotionInstructionActive := FALSE;
	END_IF
END_IF

// set outputs
//q_lrPosition
IF fbHomeIn.q_xActive THEN
	q_lrPosition := fbHomeIn.q_lrPosition;
ELSIF fbHomeTP.q_xActive THEN
	q_lrPosition := fbHomeTP.q_lrPosition;
ELSIF fbHomeLS.q_xActive THEN
	q_lrPosition := fbHomeLS.q_lrPosition;
ELSIF fbHomeTorque.q_xActive THEN
	q_lrPosition := fbHomeTorque.q_lrPosition;
ELSIF fbVarioPosJerk.q_xActive OR xDetectSetPosHomeOnPos THEN
	q_lrPosition           := lrPositionOpmMoveOnPos;
	xDetectSetPosHomeOnPos := FALSE;
ELSIF fbHomeAbs.q_xActive THEN
	q_lrPosition := fbHomeAbs.q_lrPosition;
ELSIF fbSetPos.q_xActive THEN
	q_lrPosition := fbSetPos.q_lrPosition;
ELSIF i_ifDrive <> 0 AND i_xEnable THEN
	q_lrPosition := i_ifDrive.lrPosition;
END_IF
// q_lrEncoderPosition
IF fbSetPos.i_xEnable AND fbSetPos.q_xActive THEN
	q_lrEncoderPosition := fbSetPos.q_lrEncoderPosition;
ELSIF THIS^.stSetPos_loc.iq_lencAxis <> 0 THEN
	q_lrEncoderPosition := THIS^.stSetPos_loc.iq_lencAxis.lrPosition;
ELSE
	q_lrEncoderPosition := 0.0;
END_IF

(* ---- PDL_FB_HomeAbs.fb.st ---- *)
FUNCTION_BLOCK PDL_FB_HomeAbs
VAR_INPUT
	i_xEnable        : BOOL;
	i_ifDrive        : MOIN.IF_Axis;
	i_lrHomePosition : LREAL;
	i_lrAbsEncOffset : LREAL;
	i_lrUserPeriod   : LREAL;
	i_xExecute       : BOOL;
END_VAR
VAR_OUTPUT
	q_xActive       : BOOL;
	q_xReady        : BOOL;
	q_xBusy         : BOOL;
	q_xDone         : BOOL;
	q_etDiag        : GD.ET_Diag     := GD.ET_Diag.Ok;
	q_etDiagExt     : PDL_ET_DiagExt := PDL_ET_DiagExt.Disabled;
	q_sMsg          : STRING[80];
	q_xDisableDrive : BOOL;
	q_lrPosition    : LREAL;
	q_xHomeOk       : BOOL;
END_VAR
VAR
	xEnableFlag      : BOOL;
	diState          : DINT;
	lrEncoderPeriode : LREAL;
	lrSavePosition   : LREAL;
	fbTonTimeOut     : TON;
	lrHomePosition   : LREAL;
	lrSetPosPosition : LREAL;
	fbHomeSetPos     : PDL_FB_HomeSetpos;
	lrVelocity       : LREAL;
	fbMovingAverage  : PDL_FB_MovingAverage;
	lrTurns          : LREAL;
	diSercosState    : DINT;

	ifScalingAccess     : DMFI.IF_ScalingAccess;
	ifScaling           : DMFI.IF_Scaling;
	ifDrive2Access      : DDI.IF_Drive2Access;
	ifDrive2            : DDI.IF_Drive2;
	ifDriveAccess       : DMFI.IF_DriveAccess;
	ifDrive             : DMFI.IF_Drive;
	ifDriveConfigAccess : DDI.IF_DriveConfigAccess;
	ifDriveConfig       : DDI.IF_DriveConfig;
	ifMotorAccess       : DDI.IF_MotorAccess;
	ifMotor             : DDI.IF_Motor;
	ifEncoderAccess     : DDI.IF_EncoderAccess;
	ifEncoder           : DDI.IF_Encoder;
	ifLXM62DriveAccess  : LXM62SI.IF_Lexium62DriveAccess;
	ifLXM62Drive        : LXM62SI.IF_Lexium62Drive;
	ifDeviceType		: DeviceTypeInterfaces.IF_Device_Type;

	xInterfacesInitialized : BOOL;
	xSuccess               : BOOL;

	sDummyString : STRING[80];
	etDiagInt    : GD.ET_Diag     := GD.ET_Diag.Ok;
	etDiagExtInt : PDL_ET_DiagExt := PDL_ET_DiagExt.Ok;

	fbSetDrvEncPosGetState                     : PDL_FB_SetDrvEncPosGetState;
	fbSetDrvEncPos                             : PDL_FB_SetDrvEncPos;
	etDiag                                     : GD.ET_Diag := GD.ET_Diag.Ok;
	etDiagExt                                  : PDL_ET_DiagExt := PDL_ET_DiagExt.Disabled;
	fbLoggerPoint                              : APL.FB_LoggerPoint;
	xError                                     : BOOL;
	etResult                                   : SE_Async.ET_Result;
	sResultMsg                                 : STRING(80);
	lrQuotientEncPeriodToUserPeriod            : LREAL;
	diTruncFromQuotient                        : DINT;
	lrAbsDifferenceQuotientToTruncFromQuotient : LREAL;
	xUserPeriodFitsIntoEncoderPeriod           : BOOL;
END_VAR

VAR CONSTANT
	c_lrNoVel         : LREAL := 10.0;
	c_timDisableTime  : TIME  := T#1500MS;
	c_timProgramTime  : TIME  := T#3000MS;
	c_timSettlingTime : TIME  := T#400MS;
END_VAR

IF i_xEnable AND NOT xEnableFlag THEN (* Pos. edge on Enable *)
	xEnableFlag := TRUE;
	THIS^.fbLoggerPoint.AddLogEntry(
		i_etLogLevel := APL.ET_LogLevel.UserAction,
		i_etDiag     := q_etDiag,
		i_udiDiagExt := q_etDiagExt,
		i_sMessage   := 'enable function block',
		q_etDiag     =>,
		q_etDiagExt  =>
	);
	q_xActive       := TRUE;
	q_xReady        := FALSE;
	q_xBusy         := FALSE;
	q_xDone         := FALSE;
	q_xHomeOk       := FALSE;
	q_xDisableDrive := FALSE;
	fbTonTimeOut(IN := FALSE);
	xInterfacesInitialized := THIS^.InitInterfaces();
	IF (q_etDiag <> GD.ET_Diag.Ok) THEN
		diState := 0; // exception message is already set in ParameterCheckEnable()
	ELSE
		IF SE_Async.G_ifAsyncMgr.xInitDone THEN
			q_xReady := TRUE;
			SetDiagOutput(i_etDiag := GD.ET_Diag.Ok, i_etDiagExt := PDL_ET_DiagExt.WaitForExecute, i_sMsg := '');
			diState := 10;
		ELSE
			SE_Async.G_ifAsyncMgr.Init();
			diState := -10003;
		END_IF
	END_IF
	i_ifDrive.xIsHomed := FALSE;

ELSIF NOT i_xEnable AND xEnableFlag AND q_xActive THEN (* Neg. edge on Enable *)
	xEnableFlag := FALSE;
	THIS^.fbLoggerPoint.AddLogEntry(
		i_etLogLevel := APL.ET_LogLevel.UserAction,
		i_etDiag     := q_etDiag,
		i_udiDiagExt := q_etDiagExt,
		i_sMessage   := 'disable function block',
		q_etDiag     =>,
		q_etDiagExt  =>
	);
	fbTonTimeOut(IN := FALSE);
	fbHomeSetPos(i_xEnable := FALSE);
	xInterfacesInitialized := FALSE;

	q_xActive       := FALSE;
	q_xReady        := FALSE;
	q_xBusy         := FALSE;
	q_xDone         := FALSE;
	q_xDisableDrive := FALSE;
	q_lrPosition    := 0.0;
	q_xHomeOk       := FALSE;

	SetDiagOutput(i_etDiag := GD.ET_Diag.OK, i_etDiagExt := PDL_ET_DiagExt.Disabled, i_sMsg := '');
	diState := 0;
ELSIF NOT q_xActive THEN
	RETURN;
END_IF

// set position output cyclically
IF xInterfacesInitialized THEN
	lrVelocity   := i_ifDrive.RefVelocity;
	q_lrPosition := i_ifDrive.RefPosition;
	q_xBusy      := q_etDiag = GD.ET_Diag.Ok AND NOT q_xDone AND diState > 10;
ELSE
	diState  := 0;
	q_xReady := FALSE;
	RETURN;
END_IF

CASE diState OF
	-10001: (* WaitState for async jobs *)
		IF fbSetDrvEncPos.xDone = TRUE THEN
			diState := 24;
		END_IF
	-10002:
		IF fbSetDrvEncPosGetState.xDone = TRUE THEN
			diState := 31;
		END_IF
	-10003:
		SE_Async.G_ifAsyncMgr.Init(q_xError => xError, q_etResult => etResult, q_sResultMsg => sResultMsg);
		IF xError THEN
			AsyncExtDiagTranslation(i_etResult := etResult);
			diState := 0;
		ELSIF SE_Async.G_ifAsyncMgr.xInitDone THEN
			q_xReady := TRUE;
			SetDiagOutput(i_etDiag := GD.ET_Diag.Ok, i_etDiagExt := PDL_ET_DiagExt.WaitForExecute, i_sMsg := '');
			diState := 10;
		END_IF
	0:
		; (* Idle or Error *)
	10: (* Waiting for Start *)
		IF i_xExecute THEN
			THIS^.fbLoggerPoint.AddLogEntry(
				i_etLogLevel := APL.ET_LogLevel.UserAction,
				i_etDiag     := q_etDiag,
				i_udiDiagExt := q_etDiagExt,
				i_sMessage   := 'write position',
				q_etDiag     =>,
				q_etDiagExt  =>
			);
			lrEncoderPeriode 			:= ifEncoder.Revolutions
											* ifScaling.PositionResolution
											* TO_LREAL(ifScaling.GearIn) / TO_LREAL(ifScaling.GearOut)
											* TO_LREAL( ifEncoder.GearOut) / TO_LREAL(ifEncoder.GearIn);

						// Calculation if UserPeriod fits into EncoderPeriod
			IF (i_lrUserPeriod > CMT.Gc_lrZeroTolerance) AND (lrEncoderPeriode > CMT.Gc_lrZeroTolerance) THEN

				lrQuotientEncPeriodToUserPeriod					:= lrEncoderPeriode/i_lrUserPeriod;
				diTruncFromQuotient 							:= TRUNC(lrQuotientEncPeriodToUserPeriod);
				lrAbsDifferenceQuotientToTruncFromQuotient		:= ABS (lrQuotientEncPeriodToUserPeriod - TO_LREAL(diTruncFromQuotient));

				IF (lrAbsDifferenceQuotientToTruncFromQuotient < CMT.Gc_lrZeroTolerance)
				OR ((1 - lrAbsDifferenceQuotientToTruncFromQuotient < CMT.Gc_lrZeroTolerance) AND (lrAbsDifferenceQuotientToTruncFromQuotient <= 1)) THEN
					xUserPeriodFitsIntoEncoderPeriod	:= TRUE;
				ELSE
					xUserPeriodFitsIntoEncoderPeriod	:= FALSE;
				END_IF

			END_IF

			IF (i_lrUserPeriod < 0.0) THEN
				SetDiagOutput(	i_etDiag	:= GD.ET_Diag.InputParameterInvalid,
								i_etDiagExt := PDL_ET_DiagExt.UserPeriodRange,
								i_sMsg		:= '0.0 <= i_lrUserPeriod');
				diState := 0;
			ELSIF (i_lrUserPeriod < CMT.Gc_lrZeroTolerance) AND ( (i_lrAbsEncOffset < CMT.Gc_lrZeroTolerance) OR (i_lrAbsEncOffset > (lrEncoderPeriode - CMT.Gc_lrZeroTolerance)) ) THEN
				SetDiagOutput(	i_etDiag	:= GD.ET_Diag.InputParameterInvalid,
								i_etDiagExt := PDL_ET_DiagExt.AbsEncOffsetRange,
								i_sMsg		:= STANDARD.CONCAT('0.0 < i_lrAbsEncOffset <= ', SE_CTBX.FC_LrealToString(i_sFormat := '#0.00', i_lrInput := lrEncoderPeriode - CMT.Gc_lrZeroTolerance) ));
				diState := 0;
			(* Check if UserPeriode fits into EncoderPeriode. *)
			ELSIF (i_lrUserPeriod > CMT.Gc_lrZeroTolerance) AND NOT xUserPeriodFitsIntoEncoderPeriod THEN
				SetDiagOutput(	i_etDiag	:= GD.ET_Diag.InputParameterInvalid,
								i_etDiagExt := PDL_ET_DiagExt.UserPeriodRange,
								i_sMsg		:= STANDARD.CONCAT('i_lrUserPeriod has to be a divsior of ', SE_CTBX.FC_LrealToString(i_sFormat := '#0.00', i_lrInput := lrEncoderPeriode)));
				diState := 0;

			ELSE
				q_xHomeOk       := FALSE;
				lrSavePosition  := ifdrive.ActualPosition; (* Store position before axis disabling *)
				q_xDisableDrive := TRUE; (* The Enable of the axis is switched off externally  *)
				fbTonTimeOut(IN := TRUE, PT := c_timDisableTime);
				SetDiagOutput(i_etDiag := GD.ET_Diag.OK, i_etDiagExt := PDL_ET_DiagExt.WaitUntilDriveDisabled, i_sMsg := '');
				q_xBusy := TRUE;
				q_xDone := FALSE;
				diState := 20;

				fbMovingAverage.Init(i_uiOrder := Gc_uiMovingAverageMaxOrder, q_etDiag => etDiagInt, q_etDiagExt => etDiagExtInt);
				IF etDiagInt <> GD.ET_Diag.Ok THEN
					SetDiagOutput(
						i_etDiag    := GD.ET_Diag.UnexpectedProgramBehavior,
						i_etDiagExt := PDL_ET_DiagExt.UnexpectedFeedback,
						i_sMsg      := CONCAT('PDL_FB_MovingAverage.Init(): ', UDINT_TO_STRING(etDiagExtInt))
					);
					diState := 0;
				END_IF
			END_IF
		END_IF
	20: (* Waiting for axis disabled *)
		fbTonTimeOut();
		fbMovingAverage.Insert(i_lrValue := lrVelocity, q_etDiag => etDiagInt, q_etDiagExt => etDiagExtInt);
		IF etDiagInt <> GD.ET_Diag.Ok THEN
			SetDiagOutput(
				i_etDiag    := GD.ET_Diag.UnexpectedProgramBehavior,
				i_etDiagExt := PDL_ET_DiagExt.UnexpectedFeedback,
				i_sMsg      := CONCAT('PDL_FB_MovingAverage.Insert(): ', UDINT_TO_STRING(etDiagExtInt))
			);
			diState := 0;
		END_IF

		(* Timeout for disabling axis and axis is disabled and standing*)
		IF
			fbTonTimeOut.Q AND
			i_ifDrive.etAxisState <= Moin.ET_AxisState.Disabled AND
			ABS(fbMovingAverage.lrAverage) < c_lrNoVel AND
			(fbMovingAverage.uiLevel >= Gc_uiMovingAverageMaxOrder)
		THEN
			fbTonTimeOut(IN := FALSE);
			fbMovingAverage.Init(i_uiOrder := Gc_uiMovingAverageMaxOrder, q_etDiag => etDiagInt, q_etDiagExt => etDiagExtInt);
			IF etDiagInt <> GD.ET_Diag.Ok THEN
				SetDiagOutput(
					i_etDiag    := GD.ET_Diag.UnexpectedProgramBehavior,
					i_etDiagExt := PDL_ET_DiagExt.UnexpectedFeedback,
					i_sMsg      := CONCAT('PDL_FB_MovingAverage.Init(): ', UDINT_TO_STRING(etDiagExtInt))
				);
				diState := 0;
			END_IF
			diState := 22;
		END_IF

		(* Timeout for disabling axis and axis not standing *)
		IF fbTonTimeOut.Q AND ABS(fbMovingAverage.lrAverage) >= c_lrNoVel AND (fbMovingAverage.uiLevel >= Gc_uiMovingAverageMaxOrder) THEN
			fbTonTimeOut(IN := FALSE);
			fbMovingAverage.Init(i_uiOrder := Gc_uiMovingAverageMaxOrder, q_etDiag => etDiagInt, q_etDiagExt => etDiagExtInt);
			IF etDiagInt <> GD.ET_Diag.Ok THEN
				SetDiagOutput(
					i_etDiag    := GD.ET_Diag.UnexpectedProgramBehavior,
					i_etDiagExt := PDL_ET_DiagExt.UnexpectedFeedback,
					i_sMsg      := CONCAT('PDL_FB_MovingAverage.Init(): ', UDINT_TO_STRING(etDiagExtInt))
				);
				diState := 0;
			END_IF
			SetDiagOutput(i_etDiag := GD.ET_Diag.DriveConditionInvalid, i_etDiagExt := PDL_ET_DiagExt.DriveIsMoving, i_sMsg := '');
			diState := 0;

			(* Timeout for disabling axis and axis not disabled*)
		ELSIF fbTonTimeOut.Q AND i_ifDrive.etAxisState > MOIN.ET_AxisState.Disabled THEN
			fbTonTimeOut(IN := FALSE);
			fbMovingAverage.Init(i_uiOrder := Gc_uiMovingAverageMaxOrder, q_etDiag => etDiagInt, q_etDiagExt => etDiagExtInt);
			IF etDiagInt <> GD.ET_Diag.Ok THEN
				SetDiagOutput(
					i_etDiag    := GD.ET_Diag.UnexpectedProgramBehavior,
					i_etDiagExt := PDL_ET_DiagExt.UnexpectedFeedback,
					i_sMsg      := CONCAT('PDL_FB_MovingAverage.Init(): ', UDINT_TO_STRING(etDiagExtInt))
				);
				diState := 0;
			END_IF
			SetDiagOutput(i_etDiag := GD.ET_Diag.DriveConditionInvalid, i_etDiagExt := PDL_ET_DiagExt.DriveNotDisabled, i_sMsg := '');
			diState := 0;
		END_IF
	22:
		lrEncoderPeriode := ifEncoder.Revolutions * ifScaling.PositionResolution * TO_LREAL(ifScaling.GearIn) / TO_LREAL(ifScaling.GearOut);
		lrHomePosition   := lrSetPosPosition := i_lrHomePosition + ifDrive.ActualPosition - lrSavePosition;
		(* Bring lrHomePosition into Encoder period*)
		lrTurns := TRUNC_INT(lrHomePosition / lrEncoderPeriode);
		IF lrHomePosition < 0 THEN
			lrTurns := lrTurns - 1;
		END_IF
		lrHomePosition := lrHomePosition - lrTurns * lrEncoderPeriode;
		(* Write EEPROM depending on direction of motor *)
		IF ifScaling.InvertDirection = FALSE THEN (* Motor direction right *)
			IF lrHomePosition = lrEncoderPeriode THEN
				lrHomePosition := 0.0;
			END_IF
			fbSetDrvEncPos.lrPosition := lrHomePosition;
		ELSE (* Motor direction left *)
			IF (lrEncoderPeriode - lrHomePosition) = lrEncoderPeriode THEN
				fbSetDrvEncPos.lrPosition := 0.0;
			ELSE
				fbSetDrvEncPos.lrPosition := lrEncoderPeriode - lrHomePosition;
			END_IF
		END_IF

		fbSetDrvEncPos.ifDeviceType         := ifDeviceType;
		SE_Async.G_ifAsyncMgr.Start(i_ifAsync := fbSetDrvEncPos, q_etResult => etResult, q_sResultMsg => sResultMsg, q_xError => xError);
		IF xError THEN
			AsyncExtDiagTranslation(i_etResult := etResult);
			RETURN;
		ELSE
			diState := -10001;
		END_IF
	24:
		(* Check Result of writing *)
		IF fbSetDrvEncPos.diResultSetDrvEncPos = 0 THEN
			SetDiagOutput(i_etDiag := GD.ET_Diag.OK, i_etDiagExt := PDL_ET_DiagExt.WaitUntilEncoderWritten, i_sMsg := '');
			fbTonTimeOut(IN := TRUE, PT := c_timProgramTime);
			diState := 30; (* Wait for programming time over *)
		ELSIF fbSetDrvEncPos.diResultSetDrvEncPos = -3 THEN
			SetDiagOutput(
				i_etDiag := GD.ET_Diag.InputParameterInvalid, i_etDiagExt := PDL_ET_DiagExt.DriveInvalid, i_sMsg := 'Drive must not be virtual'
			);
			diState := 0;
		ELSIF fbSetDrvEncPos.diResultSetDrvEncPos = -4 THEN
			SetDiagOutput(
				i_etDiag := GD.ET_Diag.InputParameterInvalid, i_etDiagExt := PDL_ET_DiagExt.DriveInvalid, i_sMsg := 'Drive must not be deactivated'
			);
			diState := 0;
		ELSE (* Programming error *)
			SetDiagOutput(
				i_etDiag    := GD.ET_Diag.UnexpectedProgramBehavior,
				i_etDiagExt := PDL_ET_DiagExt.UnexpectedFeedback,
				i_sMsg      := CONCAT('SystemInterface.FC_DrvEncSetPosition: ', DINT_TO_STRING(fbSetDrvEncPos.diResultSetDrvEncPos))
			);
			diState := 0;
		END_IF
	30: (* Wait for programming done *)
		(*Execute after increasing cycle-time or asynchronous*)
		(* increased cycle time was set before and is still active *)
		fbSetDrvEncPosGetState.ifDeviceType := ifDeviceType;
		SE_Async.G_ifAsyncMgr.Start(i_ifAsync := fbSetDrvEncPosGetState, q_etResult => etResult, q_sResultMsg => sResultMsg, q_xError => xError);
		IF xError THEN
			AsyncExtDiagTranslation(i_etResult := etResult);
			RETURN;
		ELSE
			diState := -10002;
		END_IF
	31:
		fbTonTimeOut();
		(* Programming finished *)
		IF fbSetDrvEncPosGetState.diResultSetDrvEncGetState = 1 THEN
			diState := 30;
			RETURN;

		ELSIF fbSetDrvEncPosGetState.diResultSetDrvEncGetState = 0 THEN
			fbTonTimeOut(IN := FALSE);
			fbTonTimeOut(IN := TRUE, PT := c_timSettlingTime); (* Delay before reading *)
			SetDiagOutput(i_etDiag := GD.ET_Diag.Ok, i_etDiagExt := PDL_ET_DiagExt.WritingPositionDone, i_sMsg := '');
			diState := 40;

		ELSIF fbSetDrvEncPosGetState.diResultSetDrvEncGetState = 2 THEN
			SetDiagOutput(i_etDiag := GD.ET_Diag.DriveConditionInvalid, i_etDiagExt := PDL_ET_DiagExt.ProgrammingInvalidEEPROM, i_sMsg := '');
			diState := 0;
			fbTonTimeOut(IN := FALSE);

		ELSIF fbSetDrvEncPosGetState.diResultSetDrvEncGetState = 3 THEN
			SetDiagOutput(i_etDiag := GD.ET_Diag.DriveConditionInvalid, i_etDiagExt := PDL_ET_DiagExt.NoAccessToEEPROM, i_sMsg := '');
			diState := 0;
			fbTonTimeOut(IN := FALSE);

		ELSIF fbTonTimeOut.Q THEN
			fbTonTimeOut(IN := FALSE);
			SetDiagOutput(i_etDiag := GD.ET_Diag.UnexpectedProgramBehavior, i_etDiagExt := PDL_ET_DiagExt.EncoderWriteTimeOut, i_sMsg := '');
			diState := 0;
		END_IF
	40: (* Wait for settling time over *)
		fbTonTimeOut();
		IF fbTonTimeOut.Q THEN
			fbTonTimeOut(IN := FALSE);
			fbHomeSetPos(
				i_xEnable        := TRUE, (* Set axis positions to the same position *)
				i_xExecute       := TRUE,
				i_ifDrive        := i_ifDrive,
				i_etMode         := PDL_ET_HomeSetPosMode.RestorePosFromAxisencoder,
				i_lrAbsEncOffset := i_lrAbsEncOffset,
				i_lrUserPeriod   := i_lrUserPeriod
			);

			SetDiagOutput(i_etDiag := GD.ET_Diag.Ok, i_etDiagExt := PDL_ET_DiagExt.WaitUntilPositionSetFromEncoder, i_sMsg := '');
			diState := 50;
		END_IF
	50: (* wait for fbHomeSetPos finished *)
		fbHomeSetPos();

		IF fbHomeSetPos.q_etDiag <> GD.ET_Diag.Ok THEN
			sDummyString :=
				SE_CTBX.FC_MultiConcat(
					i_sString1 := 'FB_HomeSetpos error: ',
					i_sString2 := PDL_FC_EtDiagExtToString(i_etDiagExt := fbHomeSetPos.q_etDiagExt),
					i_sString3 := '',
					i_sString4 := ''
				);
			SetDiagOutput(i_etDiag := GD.ET_Diag.UnexpectedProgramBehavior, i_etDiagExt := PDL_ET_DiagExt.UnexpectedFeedback, i_sMsg := sDummyString);
			diState := 0;
		ELSIF NOT fbHomeSetPos.q_xBusy THEN (* Reading is finished without error *)
			q_xHomeOk := fbHomeSetPos.q_xHomeOk;
			fbHomeSetPos(i_xEnable := FALSE);
			q_xDisableDrive := FALSE; (* Enable Axis *)

			SetDiagOutput(i_etDiag := GD.ET_Diag.Ok, i_etDiagExt := PDL_ET_DiagExt.HomingDone, i_sMsg := '');
			q_xDone := TRUE;
			diState := 60;
		END_IF
	60: (* Wait for NOT Execute *)
		IF NOT i_xExecute THEN
			SetDiagOutput(i_etDiag := GD.ET_Diag.Ok, i_etDiagExt := PDL_ET_DiagExt.WaitForExecute, i_sMsg := '');
			diState := 10;
		END_IF
	ELSE
		SetDiagOutput(
			i_etDiag := GD.ET_Diag.UnexpectedProgramBehavior, i_etDiagExt := PDL_ET_DiagExt.UnknownState, i_sMsg := DINT_TO_STRING(diState)
		);
		diState := 0;
END_CASE

(* ---- PDL_FB_HomeForce.fb.st ---- *)
FUNCTION_BLOCK PDL_FB_HomeForce
VAR_INPUT
	i_xEnable					: BOOL;
	i_ifDrive					: MOIN.IF_Axis;
	i_lrMaxForce				: LREAL;
	i_diForceTime				: DINT;
	i_lrLowLimit				: LREAL;
	i_etMode					: PDL_ET_HomeForceMode;
	i_lrOffset					: LREAL;
	i_lrMaxTravel				: LREAL;
	i_lrHomePosition			: LREAL;
	i_lrVel						: LREAL;
	i_lrAcc						: LREAL;
	i_lrDec						: LREAL;
	i_lrJerk					: LREAL;
	i_xStart					: BOOL;
END_VAR
VAR_OUTPUT
	q_xActive					: BOOL;
	q_xReady					: BOOL;
	q_etDiag					: GD.ET_Diag := GD.ET_Diag.Ok;
	q_etDiagExt					: PDL_ET_DiagExt := PDL_ET_DiagExt.Disabled;
	q_sMsg						: STRING[80];
	q_xMotionInstructionActive	: BOOL;
	q_lrPosition				: LREAL;
	q_xHomeOk					: BOOL;
END_VAR
VAR

END_VAR

(* ---- PDL_FB_HomeIn.fb.st ---- *)
FUNCTION_BLOCK PDL_FB_HomeIn
VAR_INPUT
	i_xEnable         : BOOL;
	i_ifDrive         : MOIN.IF_Axis;
	i_xSensor         : BOOL;
	i_etMode          : PDL_ET_HomeInMode;
	i_lrOffset        : LREAL;
	i_lrMaxTravel     : LREAL;
	i_lrHomePosition  : LREAL;
	i_lrVel           : LREAL;
	i_lrAcc           : LREAL;
	i_lrDec           : LREAL;
	i_lrJerk          : LREAL;
	i_xHwLimitNeg     : BOOL;
	i_xHwLimitPos     : BOOL;
	i_xRotativeSystem : BOOL;
	i_xStart          : BOOL;
END_VAR
VAR_OUTPUT
	q_xActive                  : BOOL;
	q_xReady                   : BOOL;
	q_etDiag                   : GD.ET_Diag := GD.ET_Diag.Ok;
	q_etDiagExt                : PDL_ET_DiagExt := PDL_ET_DiagExt.Disabled;
	q_sMsg                     : STRING[80];
	q_xMotionInstructionActive : BOOL;
	q_lrPosition               : LREAL;
	q_xHomeOk                  : BOOL;
END_VAR
VAR
	xSuccess                 : BOOL;
	xInterfacesInitialised   : BOOL;
	xEnableFlag              : BOOL;
	diState                  : DINT;
	lrDistance               : LREAL;
	xLimitPos                : BOOL;
	xLimitNeg                : BOOL;
	xTPPosEdge               : BOOL;
	fbStartEdge              : Standard.R_TRIG;
	fbSensorNegEdge          : Standard.F_TRIG;
	fbSensorPosEdge          : Standard.R_TRIG;
	fbLoggerPoint            : APL.FB_LoggerPoint;
	xLimitChange             : BOOL;
	fbHalt                   : PLCO.MC_Halt;
	fbStop                   : PLCO.MC_Stop;
	fbMoveRelative           : PLCO.MC_MoveRelative;
	fbSetPos                 : PLCO.MC_SetPosition;
	fbPosIN                  : PDL_FB_PosIn;
	ifDriveConfigAccess      : DDI.IF_DriveConfigAccess;
	ifDriveConfig            : DDI.IF_DriveConfig;
	ifDeviceTreeObjectAccess : UFMPLCI.IF_DeviceTreeObjectAccess;
	sDriveName               : STRING(80);

END_VAR

IF i_xEnable AND NOT xEnableFlag THEN
	xEnableFlag := TRUE;
	THIS^.fbLoggerPoint.AddLogEntry(
		i_etLogLevel := APL.ET_LogLevel.UserAction,
		i_etDiag     := q_etDiag,
		i_udiDiagExt := q_etDiagExt,
		i_sMessage   := 'enable function block',
		q_etDiag     =>,
		q_etDiagExt  =>
	);
	diState                    := 0;
	q_xActive                  := TRUE;
	q_xReady                   := FALSE;
	q_xMotionInstructionActive := FALSE;
	q_xHomeOk                  := FALSE;
	SetDiagOutput(i_etDiag := GD.ET_Diag.OK, i_etDiagExt := PDL_ET_DiagExt.Initializing, i_sMsg := '');
	xSuccess := InitInterfaces();
	IF NOT xSuccess THEN
		xInterfacesInitialised := FALSE;
		RETURN;
	ELSE
		xInterfacesInitialised := TRUE;
	END_IF

	xSuccess := InputParameterCheck();
	IF NOT xSuccess THEN
		RETURN;
	END_IF
	i_ifDrive.xIsHomed         := FALSE;

	fbStartEdge(CLK := i_xStart);
	SetDiagOutput(i_etDiag := GD.ET_Diag.Ok, i_etDiagExt := PDL_ET_DiagExt.WaitForStart, i_sMsg := '');
	q_xReady := TRUE;
	diState  := 10;

ELSIF NOT i_xEnable AND xEnableFlag THEN
	xEnableFlag := FALSE;
	THIS^.fbLoggerPoint.AddLogEntry(
		i_etLogLevel := APL.ET_LogLevel.UserAction,
		i_etDiag     := q_etDiag,
		i_udiDiagExt := q_etDiagExt,
		i_sMessage   := 'disable function block',
		q_etDiag     =>,
		q_etDiagExt  =>
	);
	q_xReady := FALSE;
	IF xInterfacesInitialised THEN
		SetDiagOutput(i_etDiag := GD.ET_Diag.OK, i_etDiagExt := PDL_ET_DiagExt.WaitUntilDisabled, i_sMsg := '');
		diState := 100;
	ELSE
		q_xActive                  := FALSE;
		q_xMotionInstructionActive := FALSE;
		q_lrPosition               := 0.0;
		q_xHomeOk                  := FALSE;
		SetDiagOutput(i_etDiag := GD.ET_Diag.OK, i_etDiagExt := PDL_ET_DiagExt.Disabled, i_sMsg := '');
		diState := 0;
	END_IF
ELSIF NOT q_xActive THEN
	RETURN;
END_IF

IF xInterfacesInitialised AND q_xActive THEN
	IF i_ifDrive.etAxisState < MOIN.ET_AxisState.Standstill AND diState > 0 AND diState < 100 THEN
		q_xReady                   := FALSE;
		q_xMotionInstructionActive := FALSE;
		SetDiagOutput(
			i_etDiag    := GD.ET_Diag.DriveConditionInvalid,
			i_etDiagExt := PDL_ET_DiagExt.DriveNotReady,
			i_sMsg 		:= STANDARD.CONCAT(sDriveName,': AxisState < Standstill')
		);
		diState := 0;
	END_IF
	q_lrPosition := i_ifDrive.lrPosition;
	fbStartEdge(CLK := i_xStart);
	fbSensorNegEdge(CLK := i_xSensor);
	fbSensorPosEdge(CLK := i_xSensor);

	(* Die HW Limits werden je nach Modus ausgewertet - Sie müssen während der Fahrt abgefragt werden *)
	IF i_etMode = PDL_ET_HomeInMode.PosDirectionPosEdgeSensor OR i_etMode = PDL_ET_HomeInMode.PosDirectionNegEdgeSensor THEN (* pos. direction *)
		xLimitPos := i_xHWLimitPos;
		xLimitNeg := i_xHWLimitNeg;

		xLimitChange := FALSE;
	ELSE (* neg. direction *)
		xLimitPos := i_xHWLimitNeg;
		xLimitNeg := i_xHWLimitPos;

		xLimitChange := TRUE;
	END_IF
END_IF

CASE diState OF
	(*---------------------------------------------------------------------------------------------*)
	0: (* Error or finished *)
		(*---------------------------------------------------------------------------------------------*)
		;
		(*---------------------------------------------------------------------------------------------*)
	10: (* wait for Start *)
		(*---------------------------------------------------------------------------------------------*)
		IF fbStartEdge.Q THEN
			xSuccess := InputParameterCheck();
			IF NOT xSuccess THEN
				q_xReady := FALSE;
				diState  := 0;
				RETURN;
			END_IF

			CASE i_etMode OF (* Selection of Mode *)
				PDL_ET_HomeInMode.PosDirectionPosEdgeSensor: (* Mode 0:  pos. Direction until pos. Edge of TP + TPOffset*)
					lrDistance := ABS(i_lrMaxTravel);
					xTPPosEdge := TRUE;
				PDL_ET_HomeInMode.NegDirectionPosEdgeSensor: (* Mode 1:  neg. Direction until pos. Edge of TP + TPOffset*)
					lrDistance := -ABS(i_lrMaxTravel);
					xTPPosEdge := TRUE;
				PDL_ET_HomeInMode.NegDirectionNegEdgeSensor: (* Mode 2:  neg. Direction until neg. Edge of TP + TPOffset*)
					xTPPosEdge := FALSE;
					lrDistance := -ABS(i_lrMaxTravel);
				PDL_ET_HomeInMode.PosDirectionNegEdgeSensor: (* Mode 3:  pos. Direction until neg. Edge of TP + TPOffset*)
					xTPPosEdge := FALSE;
					lrDistance := ABS(i_lrMaxTravel);
				ELSE
					q_xReady := FALSE;
					SetDiagOutput(i_etDiag := GD.ET_Diag.InputParameterInvalid, i_etDiagExt := PDL_ET_DiagExt.UnknownMode, i_sMsg := '');
					diState := 0;
					RETURN;
			END_CASE

			q_xMotionInstructionActive := TRUE;
			q_xHomeOk                  := FALSE;
			(*check if Axis stands on Sensor  *)
			IF (i_xSensor = xTPPosEdge AND NOT i_xRotativeSystem) OR xLimitPos THEN
				THIS^.fbMoveRelative(Distance := -lrDistance, Execute := TRUE);
				SetDiagOutput(i_etDiag := GD.ET_Diag.Ok, i_etDiagExt := PDL_ET_DiagExt.WaitForNegEdgeOfSensor, i_sMsg := '');
				diState := 20;
			ELSE

				fbPosIN(
					i_ifDrive        := i_ifDrive,
					i_xSensor        := i_xSensor,
					i_xPosEdge       := xTPPosEdge,
					i_lrMaxTravel    := lrDistance,
					i_lrOffset       := i_lrOffset,
					i_lrVelocity     := i_lrVel,
					i_lrAcceleration := i_lrAcc,
					i_lrDeceleration := i_lrDec,
					i_lrJerk         := i_lrJerk,
					i_xStart         := TRUE
				);

				IF xLimitNeg THEN (* move free from neg. Limit Switch *)
					SetDiagOutput(i_etDiag := GD.ET_Diag.Ok, i_etDiagExt := PDL_ET_DiagExt.WaitUntilLimitSwitchFree, i_sMsg := '');
					diState := 35;
				ELSE
					SetDiagOutput(i_etDiag := GD.ET_Diag.Ok, i_etDiagExt := PDL_ET_DiagExt.WaitForSensorSignal, i_sMsg := '');

					diState := 40;
				END_IF

			END_IF
		END_IF

		(*---------------------------------------------------------------------------------------------*)
	20: (* vom LimitSwitch frei fahren *)
		(*---------------------------------------------------------------------------------------------*)
		THIS^.fbMoveRelative(Execute := TRUE);
		(* Wait neg. edge of RefSensor *)
		IF (xTPPosEdge AND fbSensorNegEdge.Q) OR (NOT xTPPosEdge AND fbSensorPosEdge.Q) THEN

			THIS^.fbMoveRelative(Execute := FALSE);
			THIS^.fbHalt(Execute := TRUE);

			IF THIS^.fbHalt.Error THEN
				q_xReady                   := FALSE;
				q_xMotionInstructionActive := FALSE;
				SetDiagOutput(
					i_etDiag    := GD.ET_Diag.UnexpectedProgramBehavior,
					i_etDiagExt := PDL_ET_DiagExt.UnexpectedFeedback,
					i_sMsg      := CONCAT('MC_Halt.ErrorID: ', PLCO.FC_EtResultToString(THIS^.fbHalt.ErrorID))
				);
				THIS^.fbHalt(Execute := FALSE);
				diState := 0;
			ELSE
				SetDiagOutput(i_etDiag := GD.ET_Diag.Ok, i_etDiagExt := PDL_ET_DiagExt.WaitUntilStopped, i_sMsg := '');
				diState := 30;
			END_IF

		ELSIF xLimitNeg = TRUE THEN
			q_xReady                   := FALSE;
			q_xMotionInstructionActive := FALSE;
			THIS^.fbHalt(Execute := TRUE, Deceleration := i_lrDec, Jerk := i_lrJerk, BufferMode := PLCO.MC_Buffer_Mode.Aborting);

			IF THIS^.fbHalt.Error THEN
				q_xReady                   := FALSE;
				q_xMotionInstructionActive := FALSE;
				SetDiagOutput(
					i_etDiag    := GD.ET_Diag.UnexpectedProgramBehavior,
					i_etDiagExt := PDL_ET_DiagExt.UnexpectedFeedback,
					i_sMsg      := CONCAT('MC_Halt.ErrorID: ', PLCO.FC_EtResultToString(THIS^.fbHalt.ErrorID))
				);
				THIS^.fbHalt(Execute := FALSE);
				diState := 0;
			ELSE
				SetDiagOutput(
					i_etDiag    := GD.ET_Diag.LimitReached,
					i_etDiagExt := SEL(xLimitChange, PDL_ET_DiagExt.HwLimitNegReached, PDL_ET_DiagExt.HwLimitPosReached),
					i_sMsg      := ''
				);
				diState := 50;
			END_IF

		ELSIF fbMoveRelative.Done THEN
			q_xMotionInstructionActive := FALSE;
			q_xReady                   := FALSE;
			SetDiagOutput(i_etDiag := GD.ET_Diag.HomingFailed, i_etDiagExt := PDL_ET_DiagExt.SensorNotFound, i_sMsg := 'Sensor not found');
			THIS^.fbMoveRelative(Execute := FALSE);
			diState := 0;

		ELSIF fbMoveRelative.Error THEN (* Error *)
			q_xReady                   := FALSE;
			q_xMotionInstructionActive := FALSE;

			SetDiagOutput(
				i_etDiag    := GD.ET_Diag.UnexpectedProgramBehavior,
				i_etDiagExt := PDL_ET_DiagExt.UnexpectedFeedback,
				i_sMsg      := CONCAT('MC_MoveRelative.ErrorID: ', PLCO.FC_EtResultToString(THIS^.fbMoveRelative.ErrorID))
			);
			THIS^.fbMoveRelative(Execute := FALSE);
			diState := 0;
		END_IF

		(*---------------------------------------------------------------------------------------------*)
	30: (* wait until stopped *)
		(*---------------------------------------------------------------------------------------------*)
		THIS^.fbHalt(Execute := TRUE);
		IF THIS^.fbHalt.Done THEN
			THIS^.fbHalt(Execute := FALSE);

			IF xLimitPos THEN
				q_xReady                   := FALSE;
				q_xMotionInstructionActive := FALSE;

				//select, which linit switch cause the issue
				SetDiagOutput(
					i_etDiag    := GD.ET_Diag.HomingFailed,
					i_etDiagExt := SEL(xLimitChange, PDL_ET_DiagExt.HwLimitPosStillActive, PDL_ET_DiagExt.HwLimitNegStillActive),
					i_sMsg      := ''
				);
				diState := 0;
			ELSE
				fbPosIN(
					i_ifDrive        := i_ifDrive,
					i_xSensor        := i_xSensor,
					i_xPosEdge       := xTPPosEdge,
					i_lrMaxTravel    := lrDistance,
					i_lrOffset       := i_lrOffset,
					i_lrVelocity     := i_lrVel,
					i_lrAcceleration := i_lrAcc,
					i_lrDeceleration := i_lrDec,
					i_lrJerk         := i_lrJerk,
					i_xStart         := TRUE
				);

				SetDiagOutput(i_etDiag := GD.ET_Diag.Ok, i_etDiagExt := PDL_ET_DiagExt.WaitForSensorSignal, i_sMsg := '');

				diState := 40;
			END_IF
		ELSIF fbHalt.Error THEN (* Error *)
			q_xReady                   := FALSE;
			q_xMotionInstructionActive := FALSE;

			SetDiagOutput(
				i_etDiag    := GD.ET_Diag.UnexpectedProgramBehavior,
				i_etDiagExt := PDL_ET_DiagExt.UnexpectedFeedback,
				i_sMsg      := CONCAT('MC_Halt.ErrorID: ', PLCO.FC_EtResultToString(THIS^.fbHalt.ErrorID))
			);
			THIS^.fbHalt(Execute := FALSE);
			diState := 0;
		END_IF

		(*---------------------------------------------------------------------------------------------*)
	35: (* wait neg. Limit free *)
		(*---------------------------------------------------------------------------------------------*)
		fbPosIN(i_xSensor := i_xSensor, i_xStart := FALSE);

		IF NOT xLimitNeg THEN
			SetDiagOutput(i_etDiag := GD.ET_Diag.Ok, i_etDiagExt := PDL_ET_DiagExt.WaitForSensorSignal, i_sMsg := '');

			diState := 40;

		ELSIF xLimitPos THEN (* positive HW LimitSwitch *)
			q_xReady                   := FALSE;
			q_xMotionInstructionActive := FALSE;

			THIS^.fbHalt(Execute := TRUE, Deceleration := i_lrDec, Jerk := i_lrJerk, BufferMode := PLCO.MC_Buffer_Mode.Aborting);

			IF THIS^.fbHalt.Error THEN
				q_xReady                   := FALSE;
				q_xMotionInstructionActive := FALSE;
				SetDiagOutput(
					i_etDiag    := GD.ET_Diag.UnexpectedProgramBehavior,
					i_etDiagExt := PDL_ET_DiagExt.UnexpectedFeedback,
					i_sMsg      := CONCAT('MC_Halt.ErrorID: ', PLCO.FC_EtResultToString(THIS^.fbHalt.ErrorID))
				);
				THIS^.fbHalt(Execute := FALSE);
				diState := 0;
			ELSE
				SetDiagOutput(i_etDiag := GD.ET_Diag.LimitReached, i_etDiagExt := PDL_ET_DiagExt.HwLimitPosReached, i_sMsg := '');
				diState := 50;
			END_IF

		ELSIF fbPosIN.q_xError THEN
			q_xReady                   := FALSE;
			q_xMotionInstructionActive := FALSE;
			SetDiagOutput(
				i_etDiag    := GD.ET_Diag.UnexpectedProgramBehavior,
				i_etDiagExt := PDL_ET_DiagExt.UnexpectedFeedback,
				i_sMsg      := CONCAT('FB_PosIn: ', PLCO.FC_EtResultToString(fbPosIN.q_diErrorId))
			);
			diState := 0;

		ELSIF fbPosIn.q_xSensorNotFound THEN
			q_xReady                   := FALSE;
			q_xMotionInstructionActive := FALSE;

			IF i_etMode = PDL_ET_HomeInMode.PosDirectionPosEdgeSensor OR i_etMode = PDL_ET_HomeInMode.PosDirectionNegEdgeSensor THEN
				(* pos. direction *)
				SetDiagOutput(i_etDiag := GD.ET_Diag.HomingFailed, i_etDiagExt := PDL_ET_DiagExt.HwLimitNegStillActive, i_sMsg := '');
			ELSE
				(* neg. direction *)
				SetDiagOutput(i_etDiag := GD.ET_Diag.HomingFailed, i_etDiagExt := PDL_ET_DiagExt.HwLimitPosStillActive, i_sMsg := '');
			END_IF
			diState := 0;

			//sensor reached but limit switch is still active
		ELSIF (xLimitPos OR xLimitNeg) AND fbPosIN.q_xInOk THEN
			IF i_etMode = PDL_ET_HomeInMode.PosDirectionPosEdgeSensor OR i_etMode = PDL_ET_HomeInMode.PosDirectionNegEdgeSensor THEN
				SetDiagOutput(i_etDiag := GD.ET_Diag.HomingFailed, i_etDiagExt := PDL_ET_DiagExt.HwLimitNegStillActive, i_sMsg := '');
			ELSE
				SetDiagOutput(i_etDiag := GD.ET_Diag.HomingFailed, i_etDiagExt := PDL_ET_DiagExt.HwLimitPosStillActive, i_sMsg := '');
			END_IF

			diState := 0;
		END_IF

		(*---------------------------------------------------------------------------------------------*)
	40: (* all Modis *)
		(*---------------------------------------------------------------------------------------------*)
		fbPosIN(i_xSensor := i_xSensor, i_xStart := FALSE);

		IF fbPosIN.q_xMoveToHomePosition THEN
			SetDiagOutput(i_etDiag := GD.ET_Diag.Ok, i_etDiagExt := PDL_ET_DiagExt.WaitForSensorSignal, i_sMsg := 'Offset movement in progress');
		END_IF

		IF xLimitNeg THEN
			q_xReady                   := FALSE;
			q_xMotionInstructionActive := FALSE;

			THIS^.fbHalt(Execute := TRUE);

			SetDiagOutput(
				i_etDiag    := GD.ET_Diag.LimitReached,
				i_etDiagExt := SEL(xLimitChange, PDL_ET_DiagExt.HwLimitNegReached, PDL_ET_DiagExt.HwLimitPosReached),
				i_sMsg      := ''
			);

			diState := 50;

		ELSIF xLimitPos THEN (* positive HW LimitSwitch *)

			THIS^.fbHalt(Execute := TRUE);

			IF fbPosIN.q_xMoveToHomePosition = FALSE THEN (* TP was not seen *)
				SetDiagOutput(i_etDiag := GD.ET_Diag.Ok, i_etDiagExt := PDL_ET_DiagExt.WaitUntilStopped, i_sMsg := '');
				diState := 60;
			ELSE
				q_xReady                   := FALSE;
				q_xMotionInstructionActive := FALSE;
				SetDiagOutput(i_etDiag := GD.ET_Diag.LimitReached, i_etDiagExt := PDL_ET_DiagExt.HwLimitPosReached, i_sMsg := '');
				diState := 50;
			END_IF

		ELSIF fbPosIN.q_xSensorNotFound THEN
			q_xReady                   := FALSE;
			q_xMotionInstructionActive := FALSE;
			SetDiagOutput(i_etDiag := GD.ET_Diag.HomingFailed, i_etDiagExt := PDL_ET_DiagExt.SensorNotFound, i_sMsg := 'Sensor not found');
			diState := 0;

		ELSIF fbPosIN.q_xError THEN
			q_xReady                   := FALSE;
			q_xMotionInstructionActive := FALSE;
			SetDiagOutput(
				i_etDiag    := GD.ET_Diag.UnexpectedProgramBehavior,
				i_etDiagExt := PDL_ET_DiagExt.UnexpectedFeedback,
				i_sMsg      := CONCAT('FB_PosIn: ', PLCO.FC_EtResultToString(fbStop.ErrorID))
			);
			diState := 0;

		ELSIF fbPosIN.q_xINOk THEN
			q_xHomeOk                  := TRUE;
			i_ifDrive.xIsHomed         := TRUE;
			q_xMotionInstructionActive := FALSE;
			THIS^.fbSetPos(Execute := TRUE, Position := i_lrHomePosition, Relative := FALSE);

			IF THIS^.fbSetPos.Error THEN
				q_xReady                   := FALSE;
				q_xMotionInstructionActive := FALSE;
				SetDiagOutput(
					i_etDiag    := GD.ET_Diag.UnexpectedProgramBehavior,
					i_etDiagExt := PDL_ET_DiagExt.UnexpectedFeedback,
					i_sMsg      := CONCAT('MC_SetPosition: ', PLCO.FC_EtResultToString(THIS^.fbSetPos.ErrorID))
				);

				THIS^.fbSetPos(Execute := FALSE);
				diState := 0;
			ELSE
				SetDiagOutput(i_etDiag := GD.ET_Diag.Ok, i_etDiagExt := PDL_ET_DiagExt.HomingDone, i_sMsg := '');
				THIS^.fbSetPos(Execute := FALSE);
				diState := 10;
			END_IF
		END_IF

		(*---------------------------------------------------------------------------------------------*)
	50: (* wait  until stopped after HW Limit and Error *)
		(*---------------------------------------------------------------------------------------------*)
		THIS^.fbHalt();
		IF THIS^.fbHalt.Done THEN
			THIS^.fbHalt(Execute := FALSE);
			q_xMotionInstructionActive := FALSE;
			diState                    := 0;
			fbLoggerPoint.AddLogEntry(
				i_etLogLevel := APL.ET_LogLevel.StatusMessage,
				i_etDiag     := q_etDiag,
				i_udiDiagExt := q_etDiagExt,
				i_sMessage   := 'Axis stopped',
				q_etDiag     =>,
				q_etDiagExt  =>
			);

		ELSIF THIS^.fbHalt.Error THEN
			q_xReady                   := FALSE;
			q_xMotionInstructionActive := FALSE;
			SetDiagOutput(
				i_etDiag    := GD.ET_Diag.UnexpectedProgramBehavior,
				i_etDiagExt := PDL_ET_DiagExt.UnexpectedFeedback,
				i_sMsg      := CONCAT('MC_Halt.ErrorID: ', PLCO.FC_EtResultToString(THIS^.fbHalt.ErrorID))
			);
			THIS^.fbHalt(Execute := FALSE);
			diState := 0;
		END_IF

		(*---------------------------------------------------------------------------------------------*)
	60: (* wait until stopped after HW Limit and no Error *)
		(*---------------------------------------------------------------------------------------------*)
		THIS^.fbHalt();
		IF THIS^.fbHalt.Done THEN

			THIS^.fbMoveRelative(Execute := TRUE, Distance := -lrDistance);

			SetDiagOutput(i_etDiag := GD.ET_Diag.Ok, i_etDiagExt := PDL_ET_DiagExt.WaitForNegEdgeOfSensor, i_sMsg := '');
			diState := 20;
		END_IF

		(*---------------------------------------------------------------------------------------------*)
	100: (* Wait until stopped after Disable  *)
		(*---------------------------------------------------------------------------------------------*)
		fbMoveRelative(Execute := FALSE);
		fbHalt(Execute := FALSE);

		IF
			i_ifDrive.etAxisState <> MOIN.ET_AxisState.Disabled AND
			i_ifDrive.etAxisState <> MOIN.ET_AxisState.ErrorStop AND
			i_ifDrive.etAxisState <> MOIN.ET_AxisState.Standstill AND
			i_ifDrive.etAxisState <> MOIN.ET_AxisState.Stopping
		THEN
			fbStop.Execute      := TRUE;
			fbStop.Deceleration := i_lrDec;
			fbStop.Jerk         := i_lrJerk;
		END_IF

		fbStop();

		//stopping done
		IF
			i_ifDrive.etAxisState = MOIN.ET_AxisState.Disabled OR
			i_ifDrive.etAxisState = MOIN.ET_AxisState.ErrorStop OR
			i_ifDrive.etAxisState = MOIN.ET_AxisState.Standstill OR
			fbStop.Done
		THEN
			xInterfacesInitialised := FALSE;
			fbStop(Axis := i_ifDrive, Execute := FALSE);
			q_xActive    := FALSE;
			q_xReady     := FALSE;
			q_lrPosition := 0.0;
			SetDiagOutput(i_etDiag := GD.ET_Diag.OK, i_etDiagExt := PDL_ET_DiagExt.Disabled, i_sMsg := '');

			diState := 0;
		END_IF

		//error
		IF fbStop.Error AND fbStop.ErrorId <> PLCO.ET_Result.StoppingInterrupted THEN
			q_xMotionInstructionActive := FALSE;

			SetDiagOutput(
				i_etDiag    := GD.ET_Diag.UnexpectedProgramBehavior,
				i_etDiagExt := PDL_ET_DiagExt.UnexpectedFeedback,
				i_sMsg      := CONCAT('MC_Stop.ErrorID: ', PLCO.FC_EtResultToString(fbStop.ErrorID))
			);
			fbStop(Execute := FALSE);
		END_IF
		(* Ende Case *)
	ELSE
		q_xReady                   := FALSE;
		q_xMotionInstructionActive := FALSE;

		SetDiagOutput(
			i_etDiag := GD.ET_Diag.UnexpectedProgramBehavior, i_etDiagExt := PDL_ET_DiagExt.UnknownState, i_sMsg := DINT_TO_STRING(diState)
		);
		diState := 0;
END_CASE

(* ---- PDL_FB_HomeLimitSwitch.fb.st ---- *)
FUNCTION_BLOCK PDL_FB_HomeLimitSwitch
VAR_INPUT
	i_xEnable        : BOOL;
	i_ifDrive        : MOIN.IF_Axis;
	i_etMode         : PDL_ET_HomeLimitSwitchMode;
	i_lrOffset       : LREAL;
	i_lrMaxTravel    : LREAL;
	i_lrHomePosition : LREAL;
	i_lrVel          : LREAL;
	i_lrLowVel       : LREAL;
	i_lrAcc          : LREAL;
	i_lrDec          : LREAL;
	i_lrJerk         : LREAL;
	i_xHwLimitNeg    : BOOL;
	i_xHwLimitPos    : BOOL;
	i_xStart         : BOOL;
END_VAR
VAR_OUTPUT
	q_xActive                  : BOOL;
	q_xReady                   : BOOL;
	q_etDiag                   : GD.ET_Diag := GD.ET_Diag.Ok;
	q_etDiagExt                : PDL_ET_DiagExt := PDL_ET_DiagExt.Disabled;
	q_sMsg                     : STRING[80];
	q_xMotionInstructionActive : BOOL;
	q_lrPosition               : LREAL;
	q_xHomeOk                  : BOOL;
END_VAR
VAR
	xSuccess               : BOOL;
	xInterfacesInitialised : BOOL;
	xEnableFlag            : BOOL;
	diState                : DINT;
	fbStop                 : PLCO.MC_Stop;
	fbMoveAbsolute         : PLCO.MC_MoveAbsolute;
	fbMoveRelative         : PLCO.MC_MoveRelative;
	fbSetPos               : PLCO.MC_SetPosition;
	lrDistance             : LREAL;
	xLimitPos              : BOOL;
	xLimitNeg              : BOOL;
	xStartFlag             : BOOL;
	fbLoggerPoint          : APL.FB_LoggerPoint;

	ifDriveConfigAccess	   : DDI.IF_DriveConfigAccess;
	ifDriveConfig		   : DDI.IF_DriveConfig;
	ifDeviceTreeObjectAccess      : UFMPLCI.IF_DeviceTreeObjectAccess;
	sDriveName                    : STRING(80);
END_VAR
VAR CONSTANT
END_VAR

IF i_xEnable AND NOT xEnableFlag THEN
	xEnableFlag := TRUE;
	THIS^.fbLoggerPoint.AddLogEntry(
		i_etLogLevel := APL.ET_LogLevel.UserAction,
		i_etDiag     := q_etDiag,
		i_udiDiagExt := q_etDiagExt,
		i_sMessage   := 'enable function block',
		q_etDiag     =>,
		q_etDiagExt  =>
	);
	q_xActive                  := TRUE;
	q_xReady                   := FALSE;
	q_xHomeOk                  := FALSE;
	q_xMotionInstructionActive := FALSE;
	SetDiagOutput(
		i_etDiag    := GD.ET_Diag.OK,
		i_etDiagExt := PDL_ET_DiagExt.Initializing,
		i_sMsg      := ''
	);

	xInterfacesInitialised := InitInterfaces();
	IF NOT xInterfacesInitialised THEN
		RETURN;
	END_IF

	xSuccess := InputParameterCheck();
	IF NOT xSuccess THEN
		RETURN;
	END_IF

	THIS^.fbSetPos(
		Execute  := TRUE,
		Position := 0.0,
		Relative := FALSE
	);

	IF THIS^.fbSetPos.Error THEN
		q_xReady                   := FALSE;
		q_xMotionInstructionActive := FALSE;
		SetDiagOutput(
			i_etDiag    := GD.ET_Diag.UnexpectedProgramBehavior,
			i_etDiagExt := PDL_ET_DiagExt.UnexpectedFeedback,
			i_sMsg      :=
				CONCAT(
					'MC_SetPosition: ',
					PLCO.FC_EtResultToString(THIS^.fbSetPos.ErrorID)
				)
		);

		THIS^.fbSetPos(Execute := FALSE);
		RETURN;
	END_IF

	THIS^.fbSetPos(Execute := FALSE);
	i_ifDrive.xIsHomed := FALSE;
	xStartFlag         := FALSE;
	q_xReady           := TRUE;
	SetDiagOutput(
		i_etDiag    := GD.ET_Diag.OK,
		i_etDiagExt := PDL_ET_DiagExt.WaitForStart,
		i_sMsg      := ''
	);
	diState := 10;

ELSIF NOT I_xEnable AND xEnableFlag THEN
	xEnableFlag := FALSE;
	THIS^.fbLoggerPoint.AddLogEntry(
		i_etLogLevel := APL.ET_LogLevel.UserAction,
		i_etDiag     := q_etDiag,
		i_udiDiagExt := q_etDiagExt,
		i_sMessage   := 'disable function block',
		q_etDiag     =>,
		q_etDiagExt  =>
	);
	q_xReady := FALSE;
	IF xInterfacesInitialised THEN
		SetDiagOutput(
			i_etDiag    := GD.ET_Diag.OK,
			i_etDiagExt := PDL_ET_DiagExt.WaitUntilDisabled,
			i_sMsg      := ''
		);
		diState := 100;
	ELSE
		q_xActive                  := FALSE;
		q_xMotionInstructionActive := FALSE;
		q_lrPosition               := 0.0;
		q_xHomeOk                  := FALSE;
		SetDiagOutput(
			i_etDiag    := GD.ET_Diag.OK,
			i_etDiagExt := PDL_ET_DiagExt.Disabled,
			i_sMsg      := ''
		);
		diState := 0;
	END_IF
END_IF

IF xInterfacesInitialised AND q_xActive THEN
	IF i_ifDrive.etAxisState < MOIN.ET_AxisState.Standstill AND diState > 0 AND diState < 100 THEN
		q_xReady                   := FALSE;
		q_xMotionInstructionActive := FALSE;
		SetDiagOutput(
			i_etDiag    := GD.ET_Diag.DriveConditionInvalid,
			i_etDiagExt := PDL_ET_DiagExt.DriveNotReady,
			i_sMsg 		:= STANDARD.CONCAT(sDriveName,': AxisState < Standstill')
		);
		diState := 0;
	END_IF
	q_lrPosition := i_ifDrive.lrPosition;
	(* The HW limits are evaluated depending on the mode – they must be queried while moving. *)
	IF i_etMode = PDL_ET_HomeLimitSwitchMode.PosDirectionPosEdgeHWLimitPos OR i_etMode = PDL_ET_HomeLimitSwitchMode.PosDirectionNegEdgeHWLimitPos THEN (* pos. direction *)
		xLimitPos := i_xHWLimitPos;
		xLimitNeg := i_xHWLimitNeg;
	ELSE (* neg. direction *)
		xLimitPos := i_xHWLimitNeg;
		xLimitNeg := i_xHWLimitPos;
	END_IF
	IF i_etMode = PDL_ET_HomeLimitSwitchMode.PosDirectionNegEdgeHWLimitPos OR i_etMode = PDL_ET_HomeLimitSwitchMode.NegDirectionNegEdgeHWLimitNeg THEN (* Öffner *)
		xLimitPos := NOT xLimitPos;
		xLimitNeg := NOT xLimitNeg;
	END_IF
END_IF

CASE diState OF

	0: (* Error or ready *)
		;
	10: (* Wait for Start *)
		IF i_xStart AND NOT xStartFlag THEN
			xStartFlag := TRUE;
			THIS^.fbLoggerPoint.AddLogEntry(
				i_etLogLevel := APL.ET_LogLevel.UserAction,
				i_etDiag     := q_etDiag,
				i_udiDiagExt := q_etDiagExt,
				i_sMessage   := 'start homing',
				q_etDiag     =>,
				q_etDiagExt  =>
			);
			xSuccess := InputParameterCheck();
			IF NOT xSuccess THEN
				q_xReady := FALSE;
				diState  := 0;
				RETURN;
			END_IF
			q_xHomeOk                  := FALSE;
			q_xMotionInstructionActive := TRUE;

			CASE i_etMode OF
				PDL_ET_HomeLimitSwitchMode.PosDirectionPosEdgeHWLimitPos: (* Mode 0:  pos. Direction until pos. Edge of HomeSignal + Offset*)
					lrDistance := ABS(i_lrMaxTravel);
				PDL_ET_HomeLimitSwitchMode.NegDirectionPosEdgeHWLimitNeg: (* Mode 1:  neg. Direction until pos. Edge of HomeSignal + Offset*)
					lrDistance := -ABS(i_lrMaxTravel);
				PDL_ET_HomeLimitSwitchMode.NegDirectionNegEdgeHWLimitNeg: (* Mode 2:  pos. Direction until neg. Edge of HomeSignal + Offset*)
					lrDistance := -ABS(i_lrMaxTravel);
				PDL_ET_HomeLimitSwitchMode.PosDirectionNegEdgeHWLimitPos: (* Mode 3:  neg. Direction until neg. Edge of HomeSignal + Offset*)
					lrDistance := ABS(i_lrMaxTravel);
				ELSE
					q_xReady := FALSE;
					SetDiagOutput(
						i_etDiag    := GD.ET_Diag.InputParameterInvalid,
						i_etDiagExt := PDL_ET_DiagExt.UnknownMode,
						i_sMsg      := ''
					);
					diState := 0;
					RETURN;
			END_CASE

			IF xLimitPos AND NOT xLimitNeg THEN (* Axis stands on LS *)
				THIS^.fbMoveRelative(
					Execute  := TRUE,
					Distance := -lrDistance,
					Velocity := i_lrVel
				);

				SetDiagOutput(
					i_etDiag    := GD.ET_Diag.OK,
					i_etDiagExt := PDL_ET_DiagExt.WaitUntilLimitSwitchFree,
					i_sMsg      := ''
				);
				diState := 30;

			ELSIF xLimitPos AND xLimitNeg THEN (* Axis stands on LS pos and neg *)
				q_xMotionInstructionActive := FALSE;
				diState                    := 0;
				IF
					i_etMode = PDL_ET_HomeLimitSwitchMode.PosDirectionPosEdgeHWLimitPos OR
					i_etMode = PDL_ET_HomeLimitSwitchMode.PosDirectionNegEdgeHWLimitPos
				THEN (* pos. direction *)
					q_xReady := FALSE;
					SetDiagOutput(
						i_etDiag    := GD.ET_Diag.LimitReached,
						i_etDiagExt := PDL_ET_DiagExt.HwLimitNegReached,
						i_sMsg      := ''
					);
				ELSE
					q_xReady := FALSE;

					SetDiagOutput(
						i_etDiag    := GD.ET_Diag.LimitReached,
						i_etDiagExt := PDL_ET_DiagExt.HwLimitPosReached,
						i_sMsg      := ''
					);
				END_IF
			ELSE (* LS is free *)
				THIS^.fbMoveRelative(
					Execute  := TRUE,
					Distance := lrDistance,
					Velocity := i_lrVel
				);

				SetDiagOutput(
					i_etDiag    := GD.ET_Diag.Ok,
					i_etDiagExt := PDL_ET_DiagExt.WaitForLimitSwitchVel,
					i_sMsg      := ''
				);
				diState := 20;
			END_IF

		ELSIF NOT i_xStart AND xStartFlag THEN
			xStartFlag := FALSE;
		END_IF
	20: (* go for Limitswitch *)
		THIS^.fbMoveRelative(Execute := TRUE);

		IF THIS^.fbMoveRelative.Error THEN
			q_xReady                   := FALSE;
			q_xMotionInstructionActive := FALSE;
			SetDiagOutput(
				i_etDiag    := GD.ET_Diag.UnexpectedProgramBehavior,
				i_etDiagExt := PDL_ET_DiagExt.UnexpectedFeedback,
				i_sMsg      := CONCAT('MC_MoveRelative.ErrorID: ',PLCO.FC_EtResultToString(THIS^.fbMoveRelative.ErrorID))
			);
			THIS^.fbMoveRelative(Execute := FALSE);
			diState := 0;

		ELSIF xLimitPos THEN
			THIS^.fbMoveRelative(Execute := FALSE);
			THIS^.fbMoveRelative(
				Execute  := TRUE,
				Distance := -lrDistance,
				Velocity := i_lrLowVel
			);

			SetDiagOutput(
				i_etDiag    := GD.ET_Diag.Ok,
				i_etDiagExt := PDL_ET_DiagExt.WaitUntilLimitSwitchFree,
				i_sMsg      := ''
			);
			diState := 30;

		ELSIF THIS^.fbMoveRelative.Done THEN (* MaxDistance reached  *)
			q_xReady                   := FALSE;
			q_xMotionInstructionActive := FALSE;
			SetDiagOutput(
				i_etDiag    := GD.ET_Diag.HomingFailed,
				i_etDiagExt := PDL_ET_DiagExt.SensorNotFound,
				i_sMsg      := ''
			);
			THIS^.fbMoveRelative(Execute := FALSE);
			diState := 0;
		END_IF
	30: (* Wait for LimitSwitch free *)
		THIS^.fbMoveRelative(Execute := TRUE);

		IF NOT xLimitPos THEN (* Limitswitch is free *)
			THIS^.fbMoveRelative(Execute := FALSE);
			THIS^.fbMoveRelative(
				Execute  := TRUE,
				Distance := lrDistance,
				Velocity := i_lrLowVel
			);

			SetDiagOutput(
				i_etDiag    := GD.ET_Diag.Ok,
				i_etDiagExt := PDL_ET_DiagExt.WaitForLimitSwitchLowVel,
				i_sMsg      := ''
			);
			diState := 40;

		ELSIF THIS^.fbMoveRelative.Error THEN
			q_xReady                   := FALSE;
			q_xMotionInstructionActive := FALSE;
			SetDiagOutput(
				i_etDiag    := GD.ET_Diag.UnexpectedProgramBehavior,
				i_etDiagExt := PDL_ET_DiagExt.UnexpectedFeedback,
				i_sMsg      := CONCAT('MC_MoveRelative.ErrorID: ',PLCO.FC_EtResultToString(THIS^.fbMoveRelative.ErrorID))
			);
			THIS^.fbMoveRelative(Execute := FALSE);
			diState := 0;

		ELSIF THIS^.fbMoveRelative.Done THEN (* MaxDistance reached  *)
			q_xReady                   := FALSE;
			q_xMotionInstructionActive := FALSE;
			SetDiagOutput(
				i_etDiag    := GD.ET_Diag.HomingFailed,
				i_etDiagExt := PDL_ET_DiagExt.SensorNotFound,
				i_sMsg      := ''
			);
			THIS^.fbMoveRelative(Execute := FALSE);
			diState := 0;

		ELSIF xLimitNeg THEN (* Wrong LS *)

			THIS^.fbMoveRelative(Execute := FALSE);
			THIS^.fbStop(Execute := TRUE);

			diState := 60;
			IF
				i_etMode = PDL_ET_HomeLimitSwitchMode.PosDirectionPosEdgeHWLimitPos OR
				i_etMode = PDL_ET_HomeLimitSwitchMode.PosDirectionNegEdgeHWLimitPos
			THEN (* pos. direction *)
				q_xReady := FALSE;
				SetDiagOutput(
					i_etDiag    := GD.ET_Diag.LimitReached,
					i_etDiagExt := PDL_ET_DiagExt.HwLimitNegReached,
					i_sMsg      := ''
				);
			ELSE
				q_xReady := FALSE;
				SetDiagOutput(
					i_etDiag    := GD.ET_Diag.LimitReached,
					i_etDiagExt := PDL_ET_DiagExt.HwLimitPosReached,
					i_sMsg      := ''
				);
			END_IF
		END_IF
	40: (* go for Limitswitch *)
		THIS^.fbMoveRelative(Execute := TRUE);

		IF THIS^.fbMoveRelative.Error THEN
			q_xReady                   := FALSE;
			q_xMotionInstructionActive := FALSE;
			SetDiagOutput(
				i_etDiag    := GD.ET_Diag.UnexpectedProgramBehavior,
				i_etDiagExt := PDL_ET_DiagExt.UnexpectedFeedback,
				i_sMsg      := CONCAT('MC_MoveRelative.ErrorID: ',PLCO.FC_EtResultToString(THIS^.fbMoveRelative.ErrorID))
			);
			THIS^.fbMoveRelative(Execute := FALSE);
			diState := 0;

		ELSIF xLimitPos THEN

			THIS^.fbMoveRelative(Execute := FALSE);
			i_ifDrive.xIsHomed := TRUE;
			THIS^.fbMoveAbsolute(
				Execute  := TRUE,
				Position := q_lrPosition + i_lrOffset
			);

			SetDiagOutput(
				i_etDiag    := GD.ET_Diag.Ok,
				i_etDiagExt := PDL_ET_DiagExt.WaitUntilOffsetReached,
				i_sMsg      := ''
			);
			diState := 50;

		ELSIF THIS^.fbMoveRelative.Done THEN (* MaxDistance reached  *)
			q_xReady                   := FALSE;
			q_xMotionInstructionActive := FALSE;
			SetDiagOutput(
				i_etDiag    := GD.ET_Diag.HomingFailed,
				i_etDiagExt := PDL_ET_DiagExt.SensorNotFound,
				i_sMsg      := ''
			);
			THIS^.fbMoveRelative(Execute := FALSE);
			diState := 0;
		END_IF
	50: (* Wait for Offset reached *)
		THIS^.fbMoveAbsolute(Execute := TRUE);

		IF THIS^.fbMoveAbsolute.Error THEN
			q_xReady                   := FALSE;
			q_xMotionInstructionActive := FALSE;
			SetDiagOutput(
				i_etDiag    := GD.ET_Diag.UnexpectedProgramBehavior,
				i_etDiagExt := PDL_ET_DiagExt.UnexpectedFeedback,
				i_sMsg      := CONCAT('MC_MoveAbsolute.ErrorID: ',PLCO.FC_EtResultToString(THIS^.fbMoveAbsolute.ErrorID))
			);
			THIS^.fbMoveAbsolute(Execute := FALSE);
			i_ifDrive.xIsHomed := FALSE;
			diState := 0;

		ELSIF THIS^.fbMoveAbsolute.Done THEN
			THIS^.fbMoveAbsolute(Execute := FALSE);
			q_xHomeOk                  := TRUE;
			q_xMotionInstructionActive := FALSE;
			THIS^.fbSetPos(
				Execute  := TRUE,
				Position := i_lrHomePosition,
				Relative := FALSE
			);

			IF THIS^.fbSetPos.Error THEN
				q_xReady                   := FALSE;
				q_xMotionInstructionActive := FALSE;
				SetDiagOutput(
					i_etDiag    := GD.ET_Diag.UnexpectedProgramBehavior,
					i_etDiagExt := PDL_ET_DiagExt.UnexpectedFeedback,
					i_sMsg      := CONCAT('MC_SetPosition: ', PLCO.FC_EtResultToString(THIS^.fbSetPos.ErrorID))
				);

				THIS^.fbSetPos(Execute := FALSE);
				diState := 0;
			ELSE
				SetDiagOutput(
					i_etDiag    := GD.ET_Diag.Ok,
					i_etDiagExt := PDL_ET_DiagExt.HomingDone,
					i_sMsg      := ''
				);
				diState := 10;
				THIS^.fbSetPos(Execute := FALSE);
			END_IF
		END_IF

	60: (* wait until stopped *)
		THIS^.fbStop(Execute := TRUE);
		IF THIS^.fbStop.Done THEN
			q_xMotionInstructionActive := FALSE;
			diState                    := 0;
		ELSIF THIS^.fbStop.Error THEN
			q_xReady                   := FALSE;
			q_xMotionInstructionActive := FALSE;
			SetDiagOutput(
				i_etDiag    := GD.ET_Diag.UnexpectedProgramBehavior,
				i_etDiagExt := PDL_ET_DiagExt.UnexpectedFeedback,
				i_sMsg      := CONCAT('MC_Stop.ErrorID: ',PLCO.FC_EtResultToString(THIS^.fbStop.ErrorID))
			);
			THIS^.fbStop(Execute := FALSE);
			diState := 0;
		END_IF
	100: (* Wait until stopped  *)
		THIS^.fbMoveAbsolute(Execute := FALSE);
		THIS^.fbMoveRelative(Execute := FALSE);

		IF
			i_ifDrive.etAxisState <> MOIN.ET_AxisState.Disabled AND
			i_ifDrive.etAxisState <> MOIN.ET_AxisState.ErrorStop AND
			i_ifDrive.etAxisState <> MOIN.ET_AxisState.Standstill AND
			i_ifDrive.etAxisState <> MOIN.ET_AxisState.Stopping
		THEN
			THIS^.fbStop.Execute := TRUE;
		END_IF

		THIS^.fbStop();

		//stopping done
		IF
			i_ifDrive.etAxisState = MOIN.ET_AxisState.Disabled OR
			i_ifDrive.etAxisState = MOIN.ET_AxisState.ErrorStop OR
			i_ifDrive.etAxisState = MOIN.ET_AxisState.Standstill OR
			fbStop.Done
		THEN
			xInterfacesInitialised := FALSE;
			fbStop(Execute := FALSE);
			q_xActive    := FALSE;
			q_xReady     := FALSE;
			q_lrPosition := 0.0;
			q_xHomeOk    := FALSE;
			SetDiagOutput(
				i_etDiag    := GD.ET_Diag.OK,
				i_etDiagExt := PDL_ET_DiagExt.Disabled,
				i_sMsg      := ''
			);

			diState := 0;
		END_IF

		//error
		IF fbStop.Error AND fbStop.ErrorId <> PLCO.ET_Result.StoppingInterrupted THEN
			q_xMotionInstructionActive := FALSE;

			SetDiagOutput(
				i_etDiag    := GD.ET_Diag.UnexpectedProgramBehavior,
				i_etDiagExt := PDL_ET_DiagExt.UnexpectedFeedback,
				i_sMsg      := CONCAT('MC_Stop.ErrorID: ', PLCO.FC_EtResultToString(fbStop.ErrorID))
			);
			fbStop(Execute := FALSE);
		END_IF
		(* Ende Case *)
	ELSE
		q_xReady                   := FALSE;
		q_xMotionInstructionActive := FALSE;

		SetDiagOutput(
			i_etDiag    := GD.ET_Diag.UnexpectedProgramBehavior,
			i_etDiagExt := PDL_ET_DiagExt.UnknownState,
			i_sMsg      := DINT_TO_STRING(diState)
		);
		diState := 0;
END_CASE
